FUNCTION_BLOCK "LIOLink_RF200"   // FB5200, SCL
TITLE = LIOLink_RFID / IO_LINK_RFID_1500
{ S7_Optimized_Access := 'FALSE' }
AUTHOR : SIOS
FAMILY : LIOLink
VERSION : 3.0
// IO-Link Device FB for SIMATIC RF200 to use with S7-300/400 controllers! / IO-Link Geraete FB fuer SIMATIC RFID zur Nutzung mit S7-1500!
   VAR_INPUT
      execute : Bool;   // Request to execute function / Auftrag starten (mit steigender Flanke)
      logicalAddr : DInt;   // Logical address of IO-Link master module (sub module for ET 200eco PN) / Logische EA-Adresse des IO-Link Master Moduls
      cap : Int := 227;   // Client Access Point; 0xB400 for ET 200eco PN, CM 8x IO-Link, else 0xE003 (227) / Client Access Point (CAP), Siemens IO-Link Master immer 227 dezimal
      readWrite : Bool;   // FALSE: read, TRUE: write / Lese-/Schreibzugriff: 0=Lesen, 1=Schreiben
      port : Int;   // Port of the IO-Link Master for the Device / Port des Geraetes am IO-Link Mastermodul
      directParameterPage : Bool;   // Read access on parameter page 0 / Lesen Parameter Page 0
      vendorName : Bool;   // Read vendor name / Lesen Herstellername
      vendorText : Bool;   // Read vendor text / Lesen Herstellertext
      productName : Bool;   // Read product name / Lesen Produktname
      productID : Bool;   // Read product ID / Lesen Produkt ID
      fwRevision : Bool;   // Read firmware revision / Lesen FW-Revision
      appSpecificName : Bool;   // Read/write application specific name / Lesen/Schreiben des spezifischen Applikationsnamen
      errorCount : Bool;   // Read number of errors / Lesen des Fehlerzaehlers
      eventHistory : Bool;   // Read event history / Lesen der Ereignishistorie
      readerStatus : Bool;   // Read reader status / Lesen des Reader Status
      tagStatus : Bool;   // Read tag status / Lesen des Variablenstatus
      uidHistory : Bool;   // Read UID history / Lesen des UID Historie
   END_VAR
   VAR_OUTPUT
      done : Bool;   // TRUE: Commanded functionality has been completed successfully / Gueltigkeit 0: Daten ungueltig ; 1: Daten gueltig
      busy : Bool;   // TRUE: FB is not finished and new output values can be expected / 0: Auftrag beendet 1: Auftrag in Bearbeitung
      error : Bool;   // TRUE: An error occurred during the execution of the FB / Fehler = 0: kein Fehler; 1: Funktionsabbruch mit Fehler
      status : Word;   // 16#0000 - 16#7FFF: Status of the FB, 16#8000 - 16#FFFF: Error identification / DP/ PNIO - Fehlerstatus ; ERROR = 1 - Kommunikationsfehler in Detail
      diagDeviceFB : "LIOLink_typeDiagnostics";   // Diagnostics information of LIOLink_Device / IO-Link - Fehlerstatus; ERROR = 1: IO-Link Fehler in Detail
   END_VAR
   VAR_IN_OUT
      data : "LIOLink_RF200_typeAll";   // Data area, device specific (Data Type) / Ablage der Gerätedaten, gerätespezifisch (Datentyp in DB)
   END_VAR
   VAR
      instDevice : "LIOLink_Device";
      statRecordParam : Struct   // Parameters to read/write specific records / Datensatzparameter (geraetespezifisch)
         index : Array[0..28] of Int;   // Index of data set / Datensatzindex
         subindex : Array[0..28] of Int;   // Subindex of data sets / Datensatzsubindex
         length : Array[0..28] of Int;   // Length of data set / Datensatzlänge
      END_STRUCT;
      statRecord : Array[0..231] of Byte;   // Record buffer
      statParameterPage0 AT statRecord : "LIOLink_typeParameterPage0";
      statVendorName AT statRecord : String[12];
      statVendorText AT statRecord : String[12];
      statProductName AT statRecord : String[24];
      statProductID AT statRecord : String[16];
      statFWRevision AT statRecord : String[12];
      statAppSpecName AT statRecord : String[32];
      statErrorCount AT statRecord : Word;
      statEventHistory AT statRecord : "LIOLink_RF200_typeEventHistory";
      statReaderStatus AT statRecord : "LIOLink_RF200_typeReaderStatus";
      statTagStatus AT statRecord : "LIOLink_RF200_typeTagStatus";
      statUIDHistory AT statRecord : "LIOLink_RF200_typeUIDHistory";
      statIndex : Int;   // Requested index
      statSubindex : Int;   // Requested subindex
      statRecordLen : Int;   // Length of record to be written
      statRequest : Int;   // Case of request (data set) / Aktueller Fall (anfgefragter Datensatz)
      statDoneOld : Bool;   // Last cycle's value of instDevice.done
   END_VAR
   VAR_TEMP
      tempIndex : Int;   // Loop index
      tempLen : Int;   // Length
   END_VAR
   VAR CONSTANT
      MODE_READ : Bool := FALSE;   // Mode to read data
      MODE_WRITE : Bool := TRUE;   // Mode to write data
      STATUS_IDLE : Word := 16#7000;   // Status: Idle
   END_VAR
   // statRecordParam.index[0] := 0;
   // statRecordParam.index[1] := 0;
   // statRecordParam.index[2] := 0;
   // statRecordParam.index[3] := 0;
   // statRecordParam.index[4] := 0;
   // statRecordParam.index[5] := 0;
   // statRecordParam.index[6] := 0;
   // statRecordParam.index[7] := 0;
   // statRecordParam.index[8] := 0;
   // statRecordParam.index[9] := 74;
   // statRecordParam.index[10] := 16;
   // statRecordParam.index[11] := 17;
   // statRecordParam.index[12] := 18;
   // statRecordParam.index[13] := 19;
   // statRecordParam.index[14] := 20;
   // statRecordParam.index[15] := 21;
   // statRecordParam.index[16] := 22;
   // statRecordParam.index[17] := 23;
   // statRecordParam.index[18] := 24;
   // statRecordParam.index[19] := 32;
   // statRecordParam.index[20] := 0;
   // statRecordParam.index[21] := 0;
   // statRecordParam.index[22] := 91;
   // statRecordParam.index[23] := 90;
   // statRecordParam.index[24] := 92;
   // statRecordParam.index[25] := 0;
   // statRecordParam.index[26] := 0;
   // statRecordParam.index[27] := 0;
   // statRecordParam.index[28] := 0;
   // statRecordParam.length[0] := 0;
   // statRecordParam.length[1] := 16;
   // statRecordParam.length[2] := 0;
   // statRecordParam.length[3] := 0;
   // statRecordParam.length[4] := 0;
   // statRecordParam.length[5] := 0;
   // statRecordParam.length[6] := 0;
   // statRecordParam.length[7] := 0;
   // statRecordParam.length[8] := 0;
   // statRecordParam.length[9] := 20;
   // statRecordParam.length[10] := 12;
   // statRecordParam.length[11] := 12;
   // statRecordParam.length[12] := 24;
   // statRecordParam.length[13] := 16;
   // statRecordParam.length[14] := 0;
   // statRecordParam.length[15] := 0;
   // statRecordParam.length[16] := 0;
   // statRecordParam.length[17] := 12;
   // statRecordParam.length[18] := 32;
   // statRecordParam.length[19] := 2;
   // statRecordParam.length[20] := 0;
   // statRecordParam.length[21] := 0;
   // statRecordParam.length[22] := 15;
   // statRecordParam.length[23] := 18;
   // statRecordParam.length[24] := 40;
   // statRecordParam.length[25] := 0;
   // statRecordParam.length[26] := 0;
   // statRecordParam.length[27] := 0;
   // statRecordParam.length[28] := 0;
BEGIN
   REGION BLOCK INFO HEADER
     //===============================================================================
     // Siemens / (c)Copyright 2020
     //-------------------------------------------------------------------------------
     // Title:            LIOLink_RF200
     // Function:         Capsule block to communicate with SIMATIC RF200 Readers
     // Library:          LIOLink
     // Author:           Siemens Industry Online Support
     // Tested with:      CPU 317-2 PN/DP FW 3.2
     // Engineering:      TIA Portal V16
     // Restrictions:     --
     // Requirements:     --
     //-------------------------------------------------------------------------------
     // Change log table:
     // Version  | Date       | Expert in charge       | Changes applied
     //----------|------------|------------------------|------------------------------
     // 01.00.00 | 11.04.2014 | Online Support         | First release
     // 02.00.00 | 30.03.2015 | Online Support         | Upgrade to TIA Portal V13 SP1, use function IO_LINK_DEVICE, only one function for S7-1200 and 1500
     // 02.01.00 | 23.10.2015 | Online Support         | Update to IO_LINK_DEVICE Version 3.1
     // 03.00.00 | 22.09.2020 | Online Support         | Upgraded FB "LIOLink_Device" to V4.0.0
     //===============================================================================
   END_REGION

   REGION INIT
     IF (#execute = TRUE AND #instDevice.status = #STATUS_IDLE) THEN
       // Request selector
       IF #directParameterPage THEN
         #statRequest := 1;
       ELSIF #eventHistory THEN
         #statRequest := 9;
       ELSIF #vendorName THEN
         #statRequest := 10;
       ELSIF #vendorText THEN
         #statRequest := 11;
       ELSIF #productName THEN
         #statRequest := 12;
       ELSIF #productID THEN
         #statRequest := 13;
       ELSIF #fwRevision THEN
         #statRequest := 17;
       ELSIF #appSpecificName THEN
         #statRequest := 18;
       ELSIF #errorCount THEN
         #statRequest := 19;
       ELSIF #tagStatus THEN
         #statRequest := 22;
       ELSIF #readerStatus THEN
         #statRequest := 23;
       ELSIF #uidHistory THEN
         #statRequest := 24;
       ELSE
         #statRequest := 0;
       END_IF;

       // Set request specific parameters
       #statIndex := #statRecordParam.index[#statRequest];
       #statSubindex := #statRecordParam.subindex[#statRequest];
       #statRecordLen := #statRecordParam.length[#statRequest];

       IF #readWrite = #MODE_WRITE THEN
         REGION write
           CASE #statRequest OF
             18:
               #statAppSpecName := #data.appSpecificName; // copy text into writing data
               #tempLen := LEN(#statAppSpecName); // determine length of text

               // Shift chars in array to remove String header
               FOR #tempIndex := 0 TO #tempLen - 1 DO
                 #statRecord[#tempIndex] := #statRecord[#tempIndex + 2]; // move [2] to [0], [3] to [1] ... until end of String
               END_FOR;

               // Fill remaining characters with null
               FOR #tempIndex := #tempLen TO #statRecordLen - 1 DO
                 #statRecord[#tempIndex] := CHAR_TO_BYTE('$00');
               END_FOR;
             ELSE // all other data sets are read only  
               ;
           END_CASE;
         END_REGION

       END_IF;
     END_IF;
   END_REGION

   REGION CALL
     #instDevice(execute     := #execute,
                 logicalAddr := #logicalAddr,
                 cap         := #cap,
                 readWrite   := #readWrite,
                 "port"      := #port,
                 index       := #statIndex,
                 subindex    := #statSubindex,
                 writeLen    := #statRecordLen,
                 timeout     := T#20s,
                 record      := #statRecord);
   END_REGION

   REGION READ
     // Copy data if available and valid
     IF #instDevice.done = TRUE AND #statDoneOld = FALSE AND #readWrite = #MODE_READ THEN
       IF (#statRequest >= 10 AND #statRequest <= 18) THEN // Only applies for STRING parameters (case 10..18)
         // add two to data set length for STRING parameters (max./current length)
         FOR #tempIndex := (#statRecordLen + 1) TO 2 BY -1 DO
           #statRecord[#tempIndex] := #statRecord[#tempIndex - 2];
         END_FOR; // Shift chars in array to make space for max/current length of STRING

         #statRecord[0] := INT_TO_BYTE(#statRecordLen); // manipulate array values for STRING 
         #statRecord[1] := INT_TO_BYTE(#statRecordLen);
       END_IF; // Shift all strings and add string header 

       CASE #statRequest OF
         1:
           #data.directParameterPage := #statParameterPage0;
         9:
           #data.eventHistory := #statEventHistory;
         10:
           #data.vendorName := #statVendorName;
         11:
           #data.vendorText := #statVendorText;
         12:
           #data.productName := #statProductName;
         13:
           #data.productID := #statProductID;
         17:
           #data.fwRevision := #statFWRevision;
         18:
           #data.appSpecificName := #statAppSpecName;
         19:
           #data.errorCount := #statErrorCount;
         22:
           #data.tagStatus := #statTagStatus;
         23:
           #data.readerStatus := #statReaderStatus;
         24:
           #data.uidHistory := #statUIDHistory;
         ELSE // Other data sets are not defined
           ;
       END_CASE;
     END_IF;

     #statDoneOld := #instDevice.done;
   END_REGION

   REGION OUTPUTS
     #done := #instDevice.done;
     #busy := #instDevice.busy;
     #error := #instDevice.error;
     #status := #instDevice.status;
     #diagDeviceFB := #instDevice.diagnostics;
   END_REGION
END_FUNCTION_BLOCK

// folder: Device-specific blocks/SIRIUS

FUNCTION_BLOCK "LIOLink_3RA"   // FB5100, SCL
TITLE = LIOLink_3RA / IO_LINK_3RAxy
{ S7_Optimized_Access := 'FALSE' }
AUTHOR : SIOS
FAMILY : LIOLink
VERSION : 3.0
// IO-Link Device FB for SIRIUS 3RAxy to use with S7-300/400 controllers! / IO-Link Geraete FB fuer SIRIUS 3RAxy zur Nutzung mit S7-1500!
   VAR_INPUT
      execute : Bool;   // Request to execute function / Auftrag starten (mit steigender Flanke)
      logicalAddr : DInt;   // Logical address of IO-Link master module (sub module for ET 200eco PN) / Logische EA-Adresse des IO-Link Master Moduls
      cap : Int := 227;   // Client Access Point; 0xB400 for ET 200eco PN, CM 8x IO-Link, else 0xE003 (227) / Client Access Point (CAP), Siemens IO-Link Master immer 227 dezimal
      readWrite : Bool;   // FALSE: read, TRUE: write / Lese-/Schreibzugriff: 0=Lesen, 1=Schreiben
      port : Int;   // Port of the IO-Link Master for the Device / Port des Geraetes am IO-Link Mastermodul
      parameterPage0 : Bool;   // Read access on parameter page 0 / Lesen Parameter Page 0
      parameterPage1 : Bool;   // Read/Write access on parameter page 1 / Lesen-/Schreiben Parameter Page 1
      vendorName : Bool;   // Read Vendor Name / Lesen Herstellername
      vendorText : Bool;   // Read Vendor Text / Lesen Herstellertext
      productName : Bool;   // Read Product Name / Lesen Produktname
      productID : Bool;   // Read Product ID / Lesen Produkt ID
      productText : Bool;   // Read Product Text / Lesen Produkttext
      serialNumber : Bool;   // Read Serial Number / Lesen Seriennummer
      hwRevision : Bool;   // Read HW-Revision / Lesen HW-Revision
      fwRevision : Bool;   // Read FW-Revision / Lesen FW-Revision
      appSpecificName : Bool;   // Read/Write Application Specific Name / Lesen/Schreiben des spezifischen Applikationsnamen
      diagnostics : Bool;   // Read diagnostics / Lesen der Gruppendiagnose
      actualConfig : Bool;   // Read actual configuration / Lesen der Istkonfiguration
      targetConfig : Bool;   // Read/Write target configuration / Lesen/Schreiben der Sollkonfiguration
   END_VAR
   VAR_OUTPUT
      done : Bool;   // TRUE: Commanded functionality has been completed successfully / Gueltigkeit 0: Daten ungueltig ; 1: Daten gueltig
      busy : Bool;   // TRUE: FB is not finished and new output values can be expected / 0: Auftrag beendet 1: Auftrag in Bearbeitung
      error : Bool;   // TRUE: An error occurred during the execution of the FB / Fehler = 0: kein Fehler; 1: Funktionsabbruch mit Fehler
      status : Word;   // 16#0000 - 16#7FFF: Status of the FB, 16#8000 - 16#FFFF: Error identification / DP/ PNIO - Fehlerstatus ; ERROR = 1 - Kommunikationsfehler in Detail
      diagDeviceFB : "LIOLink_typeDiagnostics";   // Diagnostics information of LIOLink_Device / IO-Link - Fehlerstatus; ERROR = 1: IO-Link Fehler in Detail
   END_VAR
   VAR_IN_OUT
      data : "LIOLink_3RA_typeAll";   // Data area, device specific (Data Type) / Ablage der Gerätedaten, gerätespezifisch (Datentyp in DB)
   END_VAR
   VAR
      instDevice : "LIOLink_Device";
      statRecordParam : Struct   // Parameters to read/write specific records / Datensatzparameter (geraetespezifisch)
         index : Array[0..28] of Int;   // Index of data set / Datensatzindex
         subindex : Array[0..28] of Int;   // Subindex of data sets / Datensatzsubindex
         length : Array[0..28] of Int;   // Length of data set / Datensatzlänge
      END_STRUCT;
      statRecord : Array[0..231] of Byte;   // Record buffer
      statParameterPage0 AT statRecord : "LIOLink_typeParameterPage0";
      statVendorName AT statRecord : String[10];
      statVendorText AT statRecord : String[58];
      statProductName AT statRecord : String[30];
      statProductID AT statRecord : String[8];
      statProductText AT statRecord : String[2];
      statSerialNumber AT statRecord : String[8];
      statHWRevision AT statRecord : String[4];
      statFWRevision AT statRecord : String[4];
      statAppSpecName AT statRecord : String[32];
      statDiagnostics AT statRecord : "DIAG_3RAxy";
      statActualConfig AT statRecord : "PARA_3RAxy";
      statTargetConfig AT statRecord : "PARA_3RAxy";
      statParameterPage1 AT statRecord : "ParameterPage1_3RAxy";
      statIndex : Int;   // Requested index
      statSubindex : Int;   // Requested subindex
      statRecordLen : Int;   // Length of record to be written
      statRequest : Int;   // Case of request (data set) / Aktueller Fall (anfgefragter Datensatz)
      statDoneOld : Bool;   // Last cycle's value of instDevice.done
   END_VAR
   VAR_TEMP
      tempIndex : Int;   // Loop index
      tempLen : Int;   // Length
   END_VAR
   VAR CONSTANT
      MODE_READ : Bool := FALSE;   // Mode to read data
      MODE_WRITE : Bool := TRUE;   // Mode to write data
      STATUS_IDLE : Word := 16#7000;   // Status: Idle
   END_VAR
   // statRecordParam.index[4] := 0;
   // statRecordParam.index[3] := 0;
   // statRecordParam.index[2] := 1;
   // statRecordParam.index[1] := 0;
   // statRecordParam.index[25] := 0;
   // statRecordParam.index[24] := 0;
   // statRecordParam.index[23] := 90;
   // statRecordParam.index[21] := 0;
   // statRecordParam.index[20] := 0;
   // statRecordParam.index[18] := 24;
   // statRecordParam.index[17] := 23;
   // statRecordParam.index[16] := 22;
   // statRecordParam.index[15] := 21;
   // statRecordParam.index[14] := 20;
   // statRecordParam.index[13] := 19;
   // statRecordParam.index[12] := 18;
   // statRecordParam.index[11] := 17;
   // statRecordParam.index[10] := 16;
   // statRecordParam.index[8] := 0;
   // statRecordParam.index[7] := 0;
   // statRecordParam.index[6] := 0;
   // statRecordParam.index[5] := 0;
   // statRecordParam.length[28] := 0;
   // statRecordParam.length[27] := 43;
   // statRecordParam.length[26] := 43;
   // statRecordParam.length[25] := 0;
   // statRecordParam.length[24] := 0;
   // statRecordParam.length[23] := 53;
   // statRecordParam.length[22] := 0;
   // statRecordParam.length[21] := 0;
   // statRecordParam.length[20] := 0;
   // statRecordParam.length[19] := 0;
   // statRecordParam.length[18] := 32;
   // statRecordParam.length[17] := 4;
   // statRecordParam.length[16] := 4;
   // statRecordParam.length[15] := 8;
   // statRecordParam.length[14] := 2;
   // statRecordParam.length[13] := 8;
   // statRecordParam.length[12] := 30;
   // statRecordParam.length[11] := 58;
   // statRecordParam.length[10] := 10;
   // statRecordParam.length[9] := 0;
   // statRecordParam.length[8] := 0;
   // statRecordParam.length[7] := 0;
   // statRecordParam.length[6] := 0;
   // statRecordParam.length[5] := 0;
   // statRecordParam.length[4] := 0;
   // statRecordParam.length[3] := 0;
   // statRecordParam.length[2] := 16;
   // statRecordParam.length[1] := 16;
   // statRecordParam.length[0] := 0;
   // statRecordParam.index[28] := 0;
   // statRecordParam.index[27] := 130;
   // statRecordParam.index[26] := 105;
BEGIN
   REGION BLOCK INFO HEADER
     //===============================================================================
     // Siemens / (c)Copyright 2020
     //-------------------------------------------------------------------------------
     // Title:            LIOLink_3RA
     // Function:         Capsule block to communicate with 3RA devices
     // Library:          LIOLink
     // Author:           Siemens Industry Online Support
     // Tested with:      CPU 317-2 PN/DP FW 3.2
     // Engineering:      TIA Portal V16
     // Restrictions:     --
     // Requirements:     --
     //-------------------------------------------------------------------------------
     // Change log table:
     // Version  | Date       | Expert in charge       | Changes applied
     //----------|------------|------------------------|------------------------------
     // 01.00.00 | 11.04.2014 | Online Support         | First release
     // 02.00.00 | 30.03.2015 | Online Support         | Upgrade to TIA Portal V13 SP1, use function IO_LINK_DEVICE, only one function for S7-1200 and 1500
     // 02.01.00 | 23.10.2015 | Online Support         | Update to IO_LINK_DEVICE V3.1.0
     // 03.00.00 | 22.09.2020 | Online Support         | Rewrote block for FB "LIOLink_Device" V4.0.0
     //===============================================================================
   END_REGION

   REGION INIT
     IF (#execute = TRUE AND #instDevice.status = #STATUS_IDLE) THEN
       // Request selector
       IF #parameterPage0 THEN
         #statRequest := 1;
       ELSIF #parameterPage1 THEN
         #statRequest := 2;
       ELSIF #vendorName THEN
         #statRequest := 10;
       ELSIF #vendorText THEN
         #statRequest := 11;
       ELSIF #productName THEN
         #statRequest := 12;
       ELSIF #productID THEN
         #statRequest := 13;
       ELSIF #productText THEN
         #statRequest := 14;
       ELSIF #serialNumber THEN
         #statRequest := 15;
       ELSIF #hwRevision THEN
         #statRequest := 16;
       ELSIF #fwRevision THEN
         #statRequest := 17;
       ELSIF #appSpecificName THEN
         #statRequest := 18;
       ELSIF #diagnostics THEN
         #statRequest := 23;
       ELSIF #actualConfig THEN
         #statRequest := 26;
       ELSIF #targetConfig THEN
         #statRequest := 27;
       ELSE
         #statRequest := 0;
       END_IF;

       #statIndex := #statRecordParam.index[#statRequest];
       #statSubindex := #statRecordParam.subindex[#statRequest];
       #statRecordLen := #statRecordParam.length[#statRequest];

       IF #readWrite = #MODE_WRITE THEN
         REGION write
           CASE #statRequest OF
             2:
               #statParameterPage1 := #data.parameterPage1;
             18:
               #statAppSpecName := #data.appSpecificName; // copy text into writing data
               #tempLen := LEN(#statAppSpecName); // determine length of text

               // Shift chars in array to remove String header
               FOR #tempIndex := 0 TO #tempLen - 1 DO
                 #statRecord[#tempIndex] := #statRecord[#tempIndex + 2]; // move [2] to [0], [3] to [1] ... until end of String
               END_FOR;

               // Fill remaining characters with null
               FOR #tempIndex := #tempLen TO #statRecordLen - 1 DO
                 #statRecord[#tempIndex] := CHAR_TO_BYTE('$00');
               END_FOR;
             27:
               #statTargetConfig := #data.targetConfig;
             ELSE // all other data sets are read only  
               ;
           END_CASE;
         END_REGION

       END_IF;
     END_IF;
   END_REGION

   REGION CALL
     #instDevice(execute     := #execute,
                 logicalAddr := #logicalAddr,
                 cap         := #cap,
                 readWrite   := #readWrite,
                 "port"      := #port,
                 index       := #statIndex,
                 subindex    := #statSubindex,
                 writeLen    := #statRecordLen,
                 timeout     := T#20s,
                 record      := #statRecord);
   END_REGION

   REGION READ
     // Copy data if available and valid
     IF #instDevice.done = TRUE AND #statDoneOld = FALSE AND #readWrite = #MODE_READ THEN
       IF (#statRequest >= 10 AND #statRequest <= 18) THEN // Only applies for STRING parameters (case 10..18)
         // add two to data set length for STRING parameters (max./current length)
         FOR #tempIndex := (#statRecordLen + 1) TO 2 BY -1 DO
           #statRecord[#tempIndex] := #statRecord[#tempIndex - 2];
         END_FOR; // Shift chars in array to make space for max/current length of STRING

         #statRecord[0] := INT_TO_BYTE(#statRecordLen); // manipulate array values for STRING 
         #statRecord[1] := INT_TO_BYTE(#statRecordLen);
       END_IF; // Shift all strings and add string header 

       CASE #statRequest OF
         1:
           #data.parameterPage0 := #statParameterPage0;
         2:
           #data.parameterPage1 := #statParameterPage1;
         10:
           #data.vendorName := #statVendorName;
         11:
           #data.vendorText := #statVendorText;
         12:
           #data.productName := #statProductName;
         13:
           #data.productID := #statProductID;
         14:
           #data.productText := #statProductText;
         15:
           #data.serialNumber := #statSerialNumber;
         16:
           #data.hwRevision := #statHWRevision;
         17:
           #data.fwRevision := #statFWRevision;
         18:
           #data.appSpecificName := #statAppSpecName;
         23:
           #data.diagnostics := #statDiagnostics;
         26:
           #data.actualConfig := #statActualConfig;
         27:
           #data.targetConfig := #statTargetConfig;
         ELSE  // all other data set are not defined
           ;
       END_CASE;
     END_IF;

     #statDoneOld := #instDevice.done;
   END_REGION

   REGION OUTPUTS
     #done := #instDevice.done;
     #busy := #instDevice.busy;
     #error := #instDevice.error;
     #status := #instDevice.status;
     #diagDeviceFB := #instDevice.diagnostics;
   END_REGION
END_FUNCTION_BLOCK

FUNCTION_BLOCK "LIOLink_3RB24"   // FB5110, SCL
TITLE = LIOLink_3RB24 / IO_LINK_3RB24_1500
{ S7_Optimized_Access := 'FALSE' }
AUTHOR : SIOS
FAMILY : LIOLink
VERSION : 3.0
// IO-Link Device FB for SIRIUS 3RB24  to use with S7-300/400 controllers! / IO-Link Geraete FB fuer SIRIUS 3RB24 zur Nutzung mit S7-1500!
   VAR_INPUT
      execute : Bool;   // Request to execute function / Auftrag starten (mit steigender Flanke)
      logicalAddr : DInt;   // Logical address of IO-Link master module (sub module for ET 200eco PN) / Logische EA-Adresse des IO-Link Master Moduls
      cap : Int := 227;   // Client Access Point; 0xB400 for ET 200eco PN, CM 8x IO-Link, else 0xE003 (227) / Client Access Point (CAP), Siemens IO-Link Master immer 227 dezimal
      readWrite : Bool;   // FALSE: read, TRUE: write / Lese-/Schreibzugriff: 0=Lesen, 1=Schreiben
      port : Int;   // Port of the IO-Link Master for the Device / Port des Geraetes am IO-Link Mastermodul
      parameterPage0 : Bool;   // Read access on parameter page 0 / Lesen Parameter Page 0
      vendorName : Bool;   // Read Vendor Name / Lesen Herstellername
      vendorText : Bool;   // Read Vendor Text / Lesen Herstellertext
      productName : Bool;   // Read product name / Lesen Produktname
      productID : Bool;   // Read product ID / Lesen Produkt ID
      productText : Bool;   // Read product text / Lesen Produkttext
      serialNumber : Bool;   // Read serial number / Lesen Seriennummer
      hwRevision : Bool;   // Read hardware revision / Lesen HW-Revision
      fwRevision : Bool;   // Read firmware revision / Lesen FW-Revision
      appSpecificName : Bool;   // Read/Write application specific name / Lesen/Schreiben des spezifischen Applikationsnamen
      processInput : Bool;   // Read process input / Lesen der Prozesseingangsdaten
      processOutput : Bool;   // Read process output / Lesen der Prozesseausgangsdaten
      diagnostics : Bool;   // Read diagnostics / Lesen der Diagnose
      measurements : Bool;   // Read measurements / Lesen der Messwerte
      presetConfigOP : Bool;   // Read/Write preset configuration operator panel / Lesen/Schreiben der Sollkonfiguration Bediengerät
      techFunctions : Bool;   // Read technology functions / Lesen der Technologiefunktionen
   END_VAR
   VAR_OUTPUT
      done : Bool;   // TRUE: Commanded functionality has been completed successfully / Gueltigkeit 0: Daten ungueltig ; 1: Daten gueltig
      busy : Bool;   // TRUE: FB is not finished and new output values can be expected / 0: Auftrag beendet 1: Auftrag in Bearbeitung
      error : Bool;   // TRUE: An error occurred during the execution of the FB / Fehler = 0: kein Fehler; 1: Funktionsabbruch mit Fehler
      status : Word;   // 16#0000 - 16#7FFF: Status of the FB, 16#8000 - 16#FFFF: Error identification / DP/ PNIO - Fehlerstatus ; ERROR = 1 - Kommunikationsfehler in Detail
      diagDeviceFB : "LIOLink_typeDiagnostics";   // Diagnostics information of LIOLink_Device / IO-Link - Fehlerstatus; ERROR = 1: IO-Link Fehler in Detail
   END_VAR
   VAR_IN_OUT
      data : "LIOLink_3RB24_typeAll";   // Data area, device specific (Data Type) / Ablage der Gerätedaten, gerätespezifisch (Datentyp in DB)
   END_VAR
   VAR
      instDevice : "LIOLink_Device";
      statRecordParam : Struct   // Parameters to read/write specific records / Datensatzparameter (geraetespezifisch)
         index : Array[0..28] of Int;   // Index of data set / Datensatzindex
         subindex : Array[0..28] of Int;   // Subindex of data sets / Datensatzsubindex
         length : Array[0..28] of Int;   // Length of data set / Datensatzlänge
      END_STRUCT;
      statRecord : Array[0..231] of Byte;   // Record buffer
      statParameterPage0 AT statRecord : "LIOLink_typeParameterPage0";
      statVendorName AT statRecord : String[10];
      statVendorText AT statRecord : String[64];
      statProductName AT statRecord : String[30];
      statProductID AT statRecord : String[12];
      statProductText AT statRecord : String[2];
      statSerialNumber AT statRecord : String[8];
      statHWRevision AT statRecord : String[4];
      statFWRevision AT statRecord : String[4];
      statAppSpecName AT statRecord : String[32];
      statDiagnostics AT statRecord : "DIAG_3RB24";
      statMeasurements AT statRecord : "MEAS_3RB24";
      statPresetConfigOP AT statRecord : "PresetConfigOP_3RB24";
      statTechFunctions AT statRecord : "TechnoFunctions_3RB24";   // Product family SIRIUS (0x60)
      statProcessInput AT statRecord : Word;
      statProcessOutput AT statRecord : Byte;
      statIndex : Int;   // Requested index
      statSubindex : Int;   // Requested subindex
      statRecordLen : Int;   // Length of record to be written
      statRequest : Int;   // Case of request (data set) / Aktueller Fall (anfgefragter Datensatz)
      statDoneOld : Bool;   // Last cycle's value of instDevice.done
   END_VAR
   VAR_TEMP
      tempIndex : Int;   // Loop index
      tempLen : Int;   // Length
   END_VAR
   VAR CONSTANT
      MODE_READ : Bool := FALSE;   // Mode to read data
      MODE_WRITE : Bool := TRUE;   // Mode to write data
      STATUS_IDLE : Word := 16#7000;   // Status: Idle
   END_VAR
   // statRecordParam.index[4] := 0;
   // statRecordParam.index[3] := 0;
   // statRecordParam.index[2] := 0;
   // statRecordParam.index[1] := 0;
   // statRecordParam.index[25] := 94;
   // statRecordParam.index[24] := 92;
   // statRecordParam.index[23] := 0;
   // statRecordParam.index[21] := 41;
   // statRecordParam.index[20] := 40;
   // statRecordParam.index[18] := 24;
   // statRecordParam.index[17] := 23;
   // statRecordParam.index[16] := 22;
   // statRecordParam.index[15] := 21;
   // statRecordParam.index[14] := 20;
   // statRecordParam.index[13] := 19;
   // statRecordParam.index[12] := 18;
   // statRecordParam.index[11] := 17;
   // statRecordParam.index[6] := 0;
   // statRecordParam.index[5] := 0;
   // statRecordParam.index[10] := 16;
   // statRecordParam.index[8] := 0;
   // statRecordParam.index[7] := 0;
   // statRecordParam.length[28] := 26;
   // statRecordParam.length[27] := 22;
   // statRecordParam.length[26] := 0;
   // statRecordParam.length[25] := 40;
   // statRecordParam.length[24] := 25;
   // statRecordParam.length[23] := 0;
   // statRecordParam.length[22] := 0;
   // statRecordParam.length[21] := 1;
   // statRecordParam.length[20] := 2;
   // statRecordParam.length[19] := 0;
   // statRecordParam.length[18] := 32;
   // statRecordParam.length[17] := 4;
   // statRecordParam.length[16] := 4;
   // statRecordParam.length[15] := 8;
   // statRecordParam.length[14] := 2;
   // statRecordParam.length[13] := 12;
   // statRecordParam.length[12] := 30;
   // statRecordParam.length[11] := 64;
   // statRecordParam.length[10] := 10;
   // statRecordParam.length[9] := 0;
   // statRecordParam.length[8] := 0;
   // statRecordParam.length[7] := 0;
   // statRecordParam.length[6] := 0;
   // statRecordParam.length[5] := 0;
   // statRecordParam.length[4] := 0;
   // statRecordParam.length[3] := 0;
   // statRecordParam.length[2] := 0;
   // statRecordParam.length[1] := 16;
   // statRecordParam.length[0] := 0;
   // statRecordParam.index[28] := 131;
   // statRecordParam.index[27] := 130;
   // statRecordParam.index[26] := 0;
BEGIN
   REGION BLOCK INFO HEADER
     //===============================================================================
     // Siemens / (c)Copyright 2020
     //-------------------------------------------------------------------------------
     // Title:            LIOLink_3RB24
     // Function:         Capsule block to communicate with 3RB24 devices
     // Library:          LIOLink
     // Author:           Siemens Industry Online Support
     // Tested with:      CPU 317-2 PN/DP FW 3.2
     // Engineering:      TIA Portal V16
     // Restrictions:     --
     // Requirements:     --
     //-------------------------------------------------------------------------------
     // Change log table:
     // Version  | Date       | Expert in charge       | Changes applied
     //----------|------------|------------------------|------------------------------
     // 01.00.00 | 11.04.2014 | Online Support         | First release
     // 02.00.00 | 30.03.2015 | Online Support         | Upgrade to TIA Portal V13 SP1, use function IO_LINK_DEVICE, only one function for S7-1200 and 1500
     // 02.01.00 | 23.10.2015 | Online Support         | Update to IO_LINK_DEVICE Version 3.1
     // 03.00.00 | 22.09.2020 | Online Support         | Rewrote block for FB "LIOLink_Device" V4.0.0
     //===============================================================================
   END_REGION

   REGION INIT
     IF (#execute = TRUE AND #instDevice.status = #STATUS_IDLE) THEN
       // Request selector
       IF #parameterPage0 THEN
         #statRequest := 1;
       ELSIF #vendorName THEN
         #statRequest := 10;
       ELSIF #vendorText THEN
         #statRequest := 11;
       ELSIF #productName THEN
         #statRequest := 12;
       ELSIF #productID THEN
         #statRequest := 13;
       ELSIF #productText THEN
         #statRequest := 14;
       ELSIF #serialNumber THEN
         #statRequest := 15;
       ELSIF #hwRevision THEN
         #statRequest := 16;
       ELSIF #fwRevision THEN
         #statRequest := 17;
       ELSIF #appSpecificName THEN
         #statRequest := 18;
       ELSIF #processInput THEN
         #statRequest := 20;
       ELSIF #processOutput THEN
         #statRequest := 21;
       ELSIF #diagnostics THEN
         #statRequest := 24;
       ELSIF #measurements THEN
         #statRequest := 25;
       ELSIF #presetConfigOP THEN
         #statRequest := 27;
       ELSIF #techFunctions THEN
         #statRequest := 28;
       ELSE
         #statRequest := 0;
       END_IF;

       // Set request specific parameters
       #statIndex := #statRecordParam.index[#statRequest];
       #statSubindex := #statRecordParam.subindex[#statRequest];
       #statRecordLen := #statRecordParam.length[#statRequest];

       IF #readWrite = #MODE_WRITE THEN
         REGION write
           CASE #statRequest OF
             18:
               #statAppSpecName := #data.appSpecificName; // copy text into writing data
               #tempLen := LEN(#statAppSpecName); // determine length of text

               // Shift chars in array to remove String header
               FOR #tempIndex := 0 TO #tempLen - 1 DO
                 #statRecord[#tempIndex] := #statRecord[#tempIndex + 2]; // move [2] to [0], [3] to [1] ... until end of String
               END_FOR;

               // Fill remaining characters with null
               FOR #tempIndex := #tempLen TO #statRecordLen - 1 DO
                 #statRecord[#tempIndex] := CHAR_TO_BYTE('$00');
               END_FOR;
             27:
               #statPresetConfigOP := #data.presetConfig;
             ELSE // all other data sets are read only  
               ;
           END_CASE;
         END_REGION

       END_IF;
     END_IF;
   END_REGION

   REGION CALL
     #instDevice(execute     := #execute,
                 logicalAddr := #logicalAddr,
                 cap         := #cap,
                 readWrite   := #readWrite,
                 "port"      := #port,
                 index       := #statIndex,
                 subindex    := #statSubindex,
                 writeLen    := #statRecordLen,
                 timeout     := T#20s,
                 record      := #statRecord);
   END_REGION

   REGION READ
     // Copy data if available and valid
     IF #instDevice.done = TRUE AND #statDoneOld = FALSE AND #readWrite = #MODE_READ THEN
       IF (#statRequest >= 10 AND #statRequest <= 18) THEN // Only applies for STRING parameters (case 10..18)
         // add two to data set length for STRING parameters (max./current length)
         FOR #tempIndex := (#statRecordLen + 1) TO 2 BY -1 DO
           #statRecord[#tempIndex] := #statRecord[#tempIndex - 2];
         END_FOR; // Shift chars in array to make space for max/current length of STRING

         #statRecord[0] := INT_TO_BYTE(#statRecordLen); // manipulate array values for STRING 
         #statRecord[1] := INT_TO_BYTE(#statRecordLen);
       END_IF; // Shift all strings and add string header 

       CASE #statRequest OF
         1:
           #data.parameterPage0 := #statParameterPage0;
         10:
           #data.vendorName := #statVendorName;
         11:
           #data.vendorText := #statVendorText;
         12:
           #data.productName := #statProductName;
         13:
           #data.productID := #statProductID;
         14:
           #data.productText := #statProductText;
         15:
           #data.serialNumber := #statSerialNumber;
         16:
           #data.hwRevision := #statHWRevision;
         17:
           #data.fwRevision := #statFWRevision;
         18:
           #data.appSpecificName := #statAppSpecName;
         20:
           #data.processInput := #statProcessInput;
         21:
           #data.processOutput := #statProcessOutput;
         24:
           #data.diagnostics := #statDiagnostics;
         25:
           #data.measuredValues := #statMeasurements;
         27:
           #data.presetConfig := #statPresetConfigOP;
         28:
           #data.techFunctions := #statTechFunctions;
         ELSE  // Other data sets are not defined
           ;
       END_CASE;
     END_IF;

     #statDoneOld := #instDevice.done;
   END_REGION

   REGION OUTPUTS
     #done := #instDevice.done;
     #busy := #instDevice.busy;
     #error := #instDevice.error;
     #status := #instDevice.status;
     #diagDeviceFB := #instDevice.diagnostics;
   END_REGION
END_FUNCTION_BLOCK

FUNCTION_BLOCK "LIOLink_3RR24"   // FB5120, SCL
TITLE = LIOLink_3RR24 / IO_LINK_3RR24_1500
{ S7_Optimized_Access := 'FALSE' }
AUTHOR : SIOS
FAMILY : LIOLink
VERSION : 3.0
// IO-Link Device FB for SIRIUS 3RR24 to use with S7-300/400 controllers! / IO-Link Geraete FB fuer SIRIUS 3RR24 zur Nutzung mit S7-1500!
   VAR_INPUT
      execute : Bool;   // Request to execute function / Auftrag starten (mit steigender Flanke)
      logicalAddr : DInt;   // Logical address of IO-Link master module (sub module for ET 200eco PN) / Logische EA-Adresse des IO-Link Master Moduls
      cap : Int := 227;   // Client Access Point; 0xB400 for ET 200eco PN, CM 8x IO-Link, else 0xE003 (227) / Client Access Point (CAP), Siemens IO-Link Master immer 227 dezimal
      readWrite : Bool;   // FALSE: read, TRUE: write / Lese-/Schreibzugriff: 0=Lesen, 1=Schreiben
      port : Int;   // Port of the IO-Link Master for the Device / Port des Geraetes am IO-Link Mastermodul
      parameterPage0 : Bool;   // Read access on parameter page 0 / Lesen Parameter Page 0
      systemCommands : Bool;   // Write system commands / Schreiben Systemkommandos
      vendorName : Bool;   // Read vendor name / Lesen Herstellername
      vendorText : Bool;   // Read vendor text / Lesen Herstellertext
      productName : Bool;   // Read product name / Lesen Produktname
      productID : Bool;   // Read product ID / Lesen Produkt ID
      serialNumber : Bool;   // Read serial number / Lesen Seriennummer
      hwRevision : Bool;   // Read hardware revision / Lesen HW-Revision
      fwRevision : Bool;   // Read firmware revision / Lesen FW-Revision
      appSpecificName : Bool;   // Read/Write application specific name / Lesen/Schreiben des spezifischen Applikationsnamen
      diagnostics : Bool;   // Read diagnostics / Lesen der Diagnose
      measurements : Bool;   // Read measurements / Lesen der Messwerte
      parameters : Bool;   // Read/Write parameters / Lesen/Schreiben der Parameter
   END_VAR
   VAR_OUTPUT
      done : Bool;   // TRUE: Commanded functionality has been completed successfully / Gueltigkeit 0: Daten ungueltig ; 1: Daten gueltig
      busy : Bool;   // TRUE: FB is not finished and new output values can be expected / 0: Auftrag beendet 1: Auftrag in Bearbeitung
      error : Bool;   // TRUE: An error occurred during the execution of the FB / Fehler = 0: kein Fehler; 1: Funktionsabbruch mit Fehler
      status : Word;   // 16#0000 - 16#7FFF: Status of the FB, 16#8000 - 16#FFFF: Error identification / DP/ PNIO - Fehlerstatus ; ERROR = 1 - Kommunikationsfehler in Detail
      diagDeviceFB : "LIOLink_typeDiagnostics";   // Diagnostics information of LIOLink_Device / IO-Link - Fehlerstatus; ERROR = 1: IO-Link Fehler in Detail
   END_VAR
   VAR_IN_OUT
      data : "LIOLink_3RR24_typeAll";   // Data area, device specific (Data Type) / Ablage der Gerätedaten, gerätespezifisch (Datentyp in DB)
   END_VAR
   VAR
      instDevice : "LIOLink_Device";
      statRecordParam : Struct   // Parameters to read/write specific records / Datensatzparameter (geraetespezifisch)
         index : Array[0..28] of Int;   // Index of data set / Datensatzindex
         subindex : Array[0..28] of Int;   // Subindex of data sets / Datensatzsubindex
         length : Array[0..28] of Int;   // Length of data set / Datensatzlänge
      END_STRUCT;
      statRecord : Array[0..231] of Byte;   // Record buffer
      statParameterPage0 AT statRecord : "LIOLink_typeParameterPage0";
      statVendorName AT statRecord : String[11];
      statVendorText AT statRecord : String[64];
      statProductName AT statRecord : String[64];
      statProductID AT statRecord : String[14];
      statSerialNumber AT statRecord : String[16];
      statHWRevision AT statRecord : String[7];
      statFWRevision AT statRecord : String[7];
      statAppSpecName AT statRecord : String[32];
      statDiagnostics AT statRecord : "DIAG_3RR24";
      statMeasurements AT statRecord : "MEAS_3RR24";
      statParameters AT statRecord : "PARA_3RR24";   // Product family SIRIUS (0x60)
      statSystemCommands AT statRecord : Byte;
      statIndex : Int;   // Requested index
      statSubindex : Int;   // Requested subindex
      statRecordLen : Int;   // Length of record to be written
      statRequest : Int;   // Case of request (data set) / Aktueller Fall (anfgefragter Datensatz)
      statDoneOld : Bool;   // Last cycle's value of instDevice.done
   END_VAR
   VAR_TEMP
      tempIndex : Int;   // Loop index
      tempLen : Int;   // Length
   END_VAR
   VAR CONSTANT
      MODE_READ : Bool := FALSE;   // Mode to read data
      MODE_WRITE : Bool := TRUE;   // Mode to write data
      STATUS_IDLE : Word := 16#7000;   // Status: Idle
   END_VAR
   // statRecordParam.index[3] := 2;
   // statRecordParam.index[2] := 0;
   // statRecordParam.index[1] := 0;
   // statRecordParam.index[0] := 0;
   // statRecordParam.index[18] := 24;
   // statRecordParam.index[17] := 23;
   // statRecordParam.index[5] := 0;
   // statRecordParam.index[4] := 0;
   // statRecordParam.index[16] := 22;
   // statRecordParam.index[15] := 21;
   // statRecordParam.index[14] := 20;
   // statRecordParam.index[13] := 19;
   // statRecordParam.index[12] := 18;
   // statRecordParam.index[11] := 17;
   // statRecordParam.index[10] := 16;
   // statRecordParam.index[9] := 0;
   // statRecordParam.index[8] := 0;
   // statRecordParam.index[7] := 0;
   // statRecordParam.index[6] := 0;
   // statRecordParam.length[28] := 62;
   // statRecordParam.length[27] := 0;
   // statRecordParam.length[26] := 0;
   // statRecordParam.length[25] := 56;
   // statRecordParam.length[24] := 30;
   // statRecordParam.length[23] := 0;
   // statRecordParam.length[22] := 0;
   // statRecordParam.length[21] := 0;
   // statRecordParam.length[20] := 0;
   // statRecordParam.length[19] := 0;
   // statRecordParam.length[18] := 32;
   // statRecordParam.length[17] := 7;
   // statRecordParam.length[16] := 7;
   // statRecordParam.length[15] := 16;
   // statRecordParam.length[14] := 0;
   // statRecordParam.length[13] := 14;
   // statRecordParam.length[12] := 64;
   // statRecordParam.length[11] := 64;
   // statRecordParam.length[10] := 11;
   // statRecordParam.length[9] := 0;
   // statRecordParam.length[8] := 0;
   // statRecordParam.length[7] := 0;
   // statRecordParam.length[6] := 0;
   // statRecordParam.length[5] := 0;
   // statRecordParam.length[4] := 0;
   // statRecordParam.length[3] := 1;
   // statRecordParam.length[2] := 0;
   // statRecordParam.length[1] := 16;
   // statRecordParam.length[0] := 0;
   // statRecordParam.index[28] := 131;
   // statRecordParam.index[27] := 0;
   // statRecordParam.index[26] := 0;
   // statRecordParam.index[25] := 94;
   // statRecordParam.index[24] := 92;
   // statRecordParam.index[23] := 0;
   // statRecordParam.index[22] := 0;
   // statRecordParam.index[21] := 0;
   // statRecordParam.index[20] := 0;
   // statRecordParam.index[19] := 0;
BEGIN
   REGION BLOCK INFO HEADER
     //===============================================================================
     // Siemens / (c)Copyright 2020
     //-------------------------------------------------------------------------------
     // Title:            LIOLink_3RR24
     // Function:         Capsule block to communicate with 3RR24 devices
     // Library:          LIOLink
     // Author:           Siemens Industry Online Support
     // Tested with:      CPU 317-2 PN/DP FW 3.2
     // Engineering:      TIA Portal V16
     // Restrictions:     --
     // Requirements:     --
     //-------------------------------------------------------------------------------
     // Change log table:
     // Version  | Date       | Expert in charge       | Changes applied
     //----------|------------|------------------------|------------------------------
     // 01.00.00 | 11.04.2014 | Online Support         | First release
     // 01.00.01 | 12.09.2014 | Online Support         | Bugfixing write case 28 (data set 131)
     // 02.00.00 | 30.03.2015 | Online Support         | Upgrade to TIA Portal V13 SP1, use function IO_LINK_DEVICE, only one function for S7-1200 and 1500
     // 02.01.00 | 23.10.2015 | Online Support         | Update to IO_LINK_DEVICE Version 3.1
     // 03.00.00 | 22.09.2020 | Online Support         | Rewrote block for FB "LIOLink_Device" V4.0.0
     //===============================================================================
   END_REGION

   REGION INIT
     IF (#execute = TRUE AND #instDevice.status = #STATUS_IDLE) THEN
       // Request selector
       IF #parameterPage0 THEN
         #statRequest := 1;
       ELSIF #systemCommands THEN
         #statRequest := 3;
       ELSIF #vendorName THEN
         #statRequest := 10;
       ELSIF #vendorText THEN
         #statRequest := 11;
       ELSIF #productName THEN
         #statRequest := 12;
       ELSIF #productID THEN
         #statRequest := 13;
       ELSIF #serialNumber THEN
         #statRequest := 15;
       ELSIF #hwRevision THEN
         #statRequest := 16;
       ELSIF #fwRevision THEN
         #statRequest := 17;
       ELSIF #appSpecificName THEN
         #statRequest := 18;
       ELSIF #diagnostics THEN
         #statRequest := 24;
       ELSIF #measurements THEN
         #statRequest := 25;
       ELSIF #parameters THEN
         #statRequest := 28;
       ELSE
         #statRequest := 0;
       END_IF;

       // Set request specific parameters
       #statIndex := #statRecordParam.index[#statRequest];
       #statSubindex := #statRecordParam.subindex[#statRequest];
       #statRecordLen := #statRecordParam.length[#statRequest];

       IF #readWrite = #MODE_WRITE THEN
         REGION write
           CASE #statRequest OF
             3:
               #statSystemCommands := #data.systemCommands;
             18:
               #statAppSpecName := #data.appSpecificName; // copy text into writing data
               #tempLen := LEN(#statAppSpecName); // determine length of text

               // Shift chars in array to remove String header
               FOR #tempIndex := 0 TO #tempLen - 1 DO
                 #statRecord[#tempIndex] := #statRecord[#tempIndex + 2]; // move [2] to [0], [3] to [1] ... until end of String
               END_FOR;

               // Fill remaining characters with null
               FOR #tempIndex := #tempLen TO #statRecordLen - 1 DO
                 #statRecord[#tempIndex] := CHAR_TO_BYTE('$00');
               END_FOR;
             28:
               #statParameters := #data.parameters;
             ELSE    // all other data set are read only
               ;
           END_CASE;
         END_REGION

       END_IF;
     END_IF;
   END_REGION

   REGION CALL
     #instDevice(execute     := #execute,
                 logicalAddr := #logicalAddr,
                 cap         := #cap,
                 readWrite   := #readWrite,
                 "port"      := #port,
                 index       := #statIndex,
                 subindex    := #statSubindex,
                 writeLen    := #statRecordLen,
                 timeout     := T#20s,
                 record      := #statRecord);
   END_REGION

   REGION READ
     // Copy data if available and valid
     IF #instDevice.done = TRUE AND #statDoneOld = FALSE AND #readWrite = #MODE_READ THEN
       IF (#statRequest >= 10 AND #statRequest <= 18) THEN // Only applies for STRING parameters (case 10..18)
         // add two to data set length for STRING parameters (max./current length)
         FOR #tempIndex := (#statRecordLen + 1) TO 2 BY -1 DO
           #statRecord[#tempIndex] := #statRecord[#tempIndex - 2];
         END_FOR; // Shift chars in array to make space for max/current length of STRING

         #statRecord[0] := INT_TO_BYTE(#statRecordLen); // manipulate array values for STRING 
         #statRecord[1] := INT_TO_BYTE(#statRecordLen);
       END_IF; // Shift all strings and add string header 

       CASE #statRequest OF
         1:
           #data.parameterPage0 := #statParameterPage0;
         10:
           #data.vendorName := #statVendorName;
         11:
           #data.vendorText := #statVendorText;
         12:
           #data.productName := #statProductName;
         13:
           #data.productID := #statProductID;
         15:
           #data.serialNumber := #statSerialNumber;
         16:
           #data.hwRevision := #statHWRevision;
         17:
           #data.fwRevision := #statFWRevision;
         18:
           #data.appSpecificName := #statAppSpecName;
         24:
           #data.diagnostics := #statDiagnostics;
         25:
           #data.measuredValues := #statMeasurements;
         28:
           #data.parameters := #statParameters;
         ELSE  // Other data sets are not defined
           ;
       END_CASE;
     END_IF;

     #statDoneOld := #instDevice.done;
   END_REGION

   REGION OUTPUTS
     #done := #instDevice.done;
     #busy := #instDevice.busy;
     #error := #instDevice.error;
     #status := #instDevice.status;
     #diagDeviceFB := #instDevice.diagnostics;
   END_REGION
END_FUNCTION_BLOCK

FUNCTION_BLOCK "LIOLink_3RS1"   // FB5130, SCL
TITLE = LIOLink_3RS1 / IO_LINK_3RS1x_1500
{ S7_Optimized_Access := 'FALSE' }
AUTHOR : SIOS
FAMILY : LIOLink
VERSION : 3.0
// Capsule block to communicate with SIRIUS 3RS1 devices with S7-300/400 Controllers / IO-Link Geraete FB fuer SIRIUS 3RS1x zur Nutzung mit S7-1500!
   VAR_INPUT
      execute : Bool;   // Request to execute function / Auftrag starten (mit steigender Flanke)
      logicalAddr : DInt;   // Logical address of IO-Link master module (sub module for ET 200eco PN) / Logische EA-Adresse des IO-Link Master Moduls
      cap : Int := 227;   // Client Access Point; 0xB400 for ET 200eco PN, CM 8x IO-Link, else 0xE003 (227) / Client Access Point (CAP), Siemens IO-Link Master immer 227 dezimal
      readWrite : Bool;   // FALSE: read, TRUE: write / Lese-/Schreibzugriff: 0=Lesen, 1=Schreiben
      port : Int;   // Port of the IO-Link Master for the Device / Port des Geraetes am IO-Link Mastermodul
      parameterPage0 : Bool;   // Read access on parameter page 0 / Lesen Parameter Page 0
      vendorName : Bool;   // Read vendor name / Lesen Herstellername
      vendorText : Bool;   // Read vendor text / Lesen Herstellertext
      productName : Bool;   // Read product name / Lesen Produktname
      productID : Bool;   // Read product ID / Lesen Produkt ID
      hwRevision : Bool;   // Read hardware revision / Lesen HW-Revision
      fwRevision : Bool;   // Read firmware revision / Lesen FW-Revision
      appSpecificName : Bool;   // Read/Write application specific name / Lesen/Schreiben des spezifischen Applikationsnamen
      diagnostics : Bool;   // Read diagnostics / Lesen der Diagnose
      measurements : Bool;   // Read measurements / Lesen der Messwerte
      parameters : Bool;   // Read/Write parameters / Lesen/Schreiben der Parameter
   END_VAR
   VAR_OUTPUT
      done : Bool;   // TRUE: Commanded functionality has been completed successfully / Gueltigkeit 0: Daten ungueltig ; 1: Daten gueltig
      busy : Bool;   // TRUE: FB is not finished and new output values can be expected / 0: Auftrag beendet 1: Auftrag in Bearbeitung
      error : Bool;   // TRUE: An error occurred during the execution of the FB / Fehler = 0: kein Fehler; 1: Funktionsabbruch mit Fehler
      status : Word;   // 16#0000 - 16#7FFF: Status of the FB, 16#8000 - 16#FFFF: Error identification / DP/ PNIO - Fehlerstatus ; ERROR = 1 - Kommunikationsfehler in Detail
      diagDeviceFB : "LIOLink_typeDiagnostics";   // Diagnostics information of LIOLink_Device / IO-Link - Fehlerstatus; ERROR = 1: IO-Link Fehler in Detail
   END_VAR
   VAR_IN_OUT
      data : "LIOLink_3RS1_typeAll";   // Data area, device specific (Data Type) / Ablage der Gerätedaten, gerätespezifisch (Datentyp in DB)
   END_VAR
   VAR
      instDevice : "LIOLink_Device";
      statRecordParam : Struct   // Parameters to read/write specific records / Datensatzparameter (geraetespezifisch)
         index : Array[0..28] of Int;   // Index of data set / Datensatzindex
         subindex : Array[0..28] of Int;   // Subindex of data sets / Datensatzsubindex
         length : Array[0..28] of Int;   // Length of data set / Datensatzlänge
      END_STRUCT;
      statRecord : Array[0..231] of Byte;   // Record buffer
      statParameterPage0 AT statRecord : "LIOLink_typeParameterPage0";
      statVendorName AT statRecord : String[11];
      statVendorText AT statRecord : String[64];
      statProductName AT statRecord : String[64];
      statProductID AT statRecord : String[14];
      statHWRevision AT statRecord : String[7];
      statFWRevision AT statRecord : String[7];
      statAppSpecName AT statRecord : String[32];
      statDiagnostics AT statRecord : "DIAG_3RS1x";
      statMeasurements AT statRecord : "MEAS_3RS1x";
      statParameters AT statRecord : "PARA_3RS1x";   // Product family SIRIUS (0x60)
      statIndex : Int;   // Requested index
      statSubindex : Int;   // Requested subindex
      statRecordLen : Int;   // Length of record to be written
      statRequest : Int;   // Case of request (data set) / Aktueller Fall (anfgefragter Datensatz)
      statDoneOld : Bool;   // Last cycle's value of instDevice.done
   END_VAR
   VAR_TEMP
      tempIndex : Int;   // Loop index
      tempLen : Int;   // Length
   END_VAR
   VAR CONSTANT
      MODE_READ : Bool := FALSE;   // Mode to read data
      MODE_WRITE : Bool := TRUE;   // Mode to write data
      STATUS_IDLE : Word := 16#7000;   // Status: Idle
   END_VAR
   // statRecordParam.index[3] := 0;
   // statRecordParam.index[2] := 0;
   // statRecordParam.index[1] := 0;
   // statRecordParam.index[0] := 0;
   // statRecordParam.index[17] := 23;
   // statRecordParam.index[16] := 22;
   // statRecordParam.index[5] := 0;
   // statRecordParam.index[4] := 0;
   // statRecordParam.index[15] := 21;
   // statRecordParam.index[14] := 20;
   // statRecordParam.index[13] := 19;
   // statRecordParam.index[12] := 18;
   // statRecordParam.index[11] := 17;
   // statRecordParam.index[10] := 16;
   // statRecordParam.index[9] := 0;
   // statRecordParam.index[8] := 0;
   // statRecordParam.index[7] := 0;
   // statRecordParam.index[6] := 0;
   // statRecordParam.length[28] := 50;
   // statRecordParam.length[27] := 0;
   // statRecordParam.length[26] := 0;
   // statRecordParam.length[25] := 46;
   // statRecordParam.length[24] := 40;
   // statRecordParam.length[23] := 0;
   // statRecordParam.length[22] := 0;
   // statRecordParam.length[21] := 0;
   // statRecordParam.length[20] := 0;
   // statRecordParam.length[19] := 0;
   // statRecordParam.length[18] := 32;
   // statRecordParam.length[17] := 7;
   // statRecordParam.length[16] := 7;
   // statRecordParam.length[15] := 0;
   // statRecordParam.length[14] := 0;
   // statRecordParam.length[13] := 14;
   // statRecordParam.length[12] := 64;
   // statRecordParam.length[11] := 64;
   // statRecordParam.length[10] := 11;
   // statRecordParam.length[9] := 0;
   // statRecordParam.length[8] := 0;
   // statRecordParam.length[7] := 0;
   // statRecordParam.length[6] := 0;
   // statRecordParam.length[5] := 0;
   // statRecordParam.length[4] := 0;
   // statRecordParam.length[3] := 0;
   // statRecordParam.length[2] := 0;
   // statRecordParam.length[1] := 16;
   // statRecordParam.length[0] := 0;
   // statRecordParam.index[28] := 131;
   // statRecordParam.index[27] := 0;
   // statRecordParam.index[26] := 0;
   // statRecordParam.index[25] := 94;
   // statRecordParam.index[24] := 92;
   // statRecordParam.index[23] := 0;
   // statRecordParam.index[22] := 0;
   // statRecordParam.index[21] := 0;
   // statRecordParam.index[20] := 0;
   // statRecordParam.index[19] := 0;
   // statRecordParam.index[18] := 24;
BEGIN
   REGION BLOCK INFO HEADER
     //===============================================================================
     // Siemens / (c)Copyright 2020
     //-------------------------------------------------------------------------------
     // Title:            LIOLink_3RS1
     // Function:         Capsule block to communicate with SIRIUS 3RS1 devices
     // Library:          LIOLink
     // Author:           Siemens Industry Online Support
     // Tested with:      CPU 317-2 PN/DP FW 3.2
     // Engineering:      TIA Portal V16
     // Restrictions:     --
     // Requirements:     --
     //-------------------------------------------------------------------------------
     // Change log table:
     // Version  | Date       | Expert in charge       | Changes applied
     //----------|------------|------------------------|------------------------------
     // 01.00.00 | 11.04.2014 | Online Support         | First release
     // 02.00.00 | 30.03.2015 | Online Support         | Upgrade to TIA Portal V13 SP1, use function IO_LINK_DEVICE, only one function for S7-1200 and 1500
     // 02.01.00 | 23.10.2015 | Online Support         | Update to IO_LINK_DEVICE Version 3.1
     // 03.00.00 | 22.09.2020 | Online Support         | Rewrote block for FB "LIOLink_Device" V4.0.0
     //===============================================================================
   END_REGION

   REGION INIT
     IF (#execute = TRUE AND #instDevice.status = #STATUS_IDLE) THEN
       // Request selector
       IF #parameterPage0 THEN
         #statRequest := 1;
       ELSIF #vendorName THEN
         #statRequest := 10;
       ELSIF #vendorText THEN
         #statRequest := 11;
       ELSIF #productName THEN
         #statRequest := 12;
       ELSIF #productID THEN
         #statRequest := 13;
       ELSIF #hwRevision THEN
         #statRequest := 16;
       ELSIF #fwRevision THEN
         #statRequest := 17;
       ELSIF #appSpecificName THEN
         #statRequest := 18;
       ELSIF #diagnostics THEN
         #statRequest := 24;
       ELSIF #measurements THEN
         #statRequest := 25;
       ELSIF #parameters THEN
         #statRequest := 28;
       ELSE
         #statRequest := 0;
       END_IF;

       // Set request specific parameters
       #statIndex := #statRecordParam.index[#statRequest];
       #statSubindex := #statRecordParam.subindex[#statRequest];
       #statRecordLen := #statRecordParam.length[#statRequest];

       IF #readWrite = #MODE_WRITE THEN
         REGION write
           CASE #statRequest OF
             18:
               #statAppSpecName := #data.appSpecificName; // copy text into writing data
               #tempLen := LEN(#statAppSpecName); // determine length of text

               // Shift chars in array to remove String header
               FOR #tempIndex := 0 TO #tempLen - 1 DO
                 #statRecord[#tempIndex] := #statRecord[#tempIndex + 2]; // move [2] to [0], [3] to [1] ... until end of String
               END_FOR;

               // Fill remaining characters with null
               FOR #tempIndex := #tempLen TO #statRecordLen - 1 DO
                 #statRecord[#tempIndex] := CHAR_TO_BYTE('$00');
               END_FOR;
             28:
               #statParameters := #data.parameters;
             ELSE // All other data sets are read only
               ;
           END_CASE;
         END_REGION

       END_IF;
     END_IF;
   END_REGION

   REGION CALL
     #instDevice(execute     := #execute,
                 logicalAddr := #logicalAddr,
                 cap         := #cap,
                 readWrite   := #readWrite,
                 "port"      := #port,
                 index       := #statIndex,
                 subindex    := #statSubindex,
                 writeLen    := #statRecordLen,
                 timeout     := T#20s,
                 record      := #statRecord);
   END_REGION

   REGION READ
     // Copy data if available and valid
     IF #instDevice.done = TRUE AND #statDoneOld = FALSE AND #readWrite = #MODE_READ THEN
       IF (#statRequest >= 10 AND #statRequest <= 18) THEN // Only applies for STRING parameters (case 10..18)
         // add two to data set length for STRING parameters (max./current length)
         FOR #tempIndex := (#statRecordLen + 1) TO 2 BY -1 DO
           #statRecord[#tempIndex] := #statRecord[#tempIndex - 2];
         END_FOR; // Shift chars in array to make space for max/current length of STRING

         #statRecord[0] := INT_TO_BYTE(#statRecordLen); // manipulate array values for STRING 
         #statRecord[1] := INT_TO_BYTE(#statRecordLen);
       END_IF; // Shift all strings and add string header 

       CASE #statRequest OF
         1:
           #data.parameterPage0 := #statParameterPage0;
         10:
           #data.vendorName := #statVendorName;
         11:
           #data.vendorText := #statVendorText;
         12:
           #data.productName := #statProductName;
         13:
           #data.productID := #statProductID;
         16:
           #data.hardwareRevision := #statHWRevision;
         17:
           #data.firmwareRevision := #statFWRevision;
         18:
           #data.appSpecificName := #statAppSpecName;
         24:
           #data.diagnostics := #statDiagnostics;
         25:
           #data.measuredValues := #statMeasurements;
         28:
           #data.parameters := #statParameters;
         ELSE  // Other data sets are not defined
           ;
       END_CASE;
     END_IF;

     #statDoneOld := #instDevice.done;
   END_REGION

   REGION OUTPUTS
     #done := #instDevice.done;
     #busy := #instDevice.busy;
     #error := #instDevice.error;
     #status := #instDevice.status;
     #diagDeviceFB := #instDevice.diagnostics;
   END_REGION
END_FUNCTION_BLOCK

FUNCTION_BLOCK "LIOLink_3RS2"   // FB5131, SCL
TITLE = LIOLink_3RS2 / IO_LINK_3RS1x_1500
{ S7_Optimized_Access := 'FALSE' }
AUTHOR : SIOS
FAMILY : LIOLink
VERSION : 1.0
// Capsule block to communicate with SIRIUS 3RS2 devices with S7-300/400 Controllers / IO-Link Geraete FB fuer SIRIUS 3RS1x zur Nutzung mit S7-1500!
   VAR_INPUT
      execute : Bool;   // Request to execute function / Auftrag starten (mit steigender Flanke)
      logicalAddr : DInt;   // Logical address of IO-Link master module (sub module for ET 200eco PN) / Logische EA-Adresse des IO-Link Master Moduls
      cap : Int := 227;   // Client Access Point; 0xB400 for ET 200eco PN, CM 8x IO-Link, else 0xE003 (227) / Client Access Point (CAP), Siemens IO-Link Master immer 227 dezimal
      readWrite : Bool;   // FALSE: read, TRUE: write / Lese-/Schreibzugriff: 0=Lesen, 1=Schreiben
      port : Int;   // Port of the IO-Link Master for the Device / Port des Geraetes am IO-Link Mastermodul
      parameterPage0 : Bool;   // Read parameter page 0 / Lesen Parameter Page 0
      vendorName : Bool;   // Read vendor name / Lesen Herstellername
      vendorText : Bool;   // Read vendor text / Lesen Herstellertext
      productName : Bool;   // Read product name / Lesen Produktname
      productID : Bool;   // Read product ID / Lesen Produkt ID
      fwRevision : Bool;   // Read firmware revision / Lesen FW-Revision
      appSpecificName : Bool;   // Read/write application specific name / Lesen/Schreiben des spezifischen Applikationsnamen
      diagnostics : Bool;   // Read diagnostics / Lesen der Diagnose
      measuredValues : Bool;   // Read measured values / Lesen der Messwerte
      parameters : Bool;   // Read/Write parameters / Lesen/Schreiben der Parameter
   END_VAR
   VAR_OUTPUT
      done : Bool;   // TRUE: Commanded functionality has been completed successfully / Gueltigkeit 0: Daten ungueltig ; 1: Daten gueltig
      busy : Bool;   // TRUE: FB is not finished and new output values can be expected / 0: Auftrag beendet 1: Auftrag in Bearbeitung
      error : Bool;   // TRUE: An error occurred during the execution of the FB / Fehler = 0: kein Fehler; 1: Funktionsabbruch mit Fehler
      status : Word;   // 16#0000 - 16#7FFF: Status of the FB, 16#8000 - 16#FFFF: Error identification / DP/ PNIO - Fehlerstatus ; ERROR = 1 - Kommunikationsfehler in Detail
      diagDeviceFB : "LIOLink_typeDiagnostics";   // Diagnostics information of LIOLink_Device / IO-Link - Fehlerstatus; ERROR = 1: IO-Link Fehler in Detail
   END_VAR
   VAR_IN_OUT
      data : "LIOLink_3RS2_typeAll";   // Data area, device specific (Data Type) / Ablage der Gerätedaten, gerätespezifisch (Datentyp in DB)
   END_VAR
   VAR
      instDevice : "LIOLink_Device";
      statRecord : Array[0..231] of Byte;   // Record buffer
      statParameterPage0 AT statRecord : "LIOLink_typeParameterPage0";
      statVendorName AT statRecord : String[11];
      statVendorText AT statRecord : String[64];
      statProductName AT statRecord : String[64];
      statProductID AT statRecord : String[14];
      statFWRevision AT statRecord : String[7];
      statAppSpecName AT statRecord : String[32];
      statDiagnostics AT statRecord : "LIOLink_3RS2_typeDiag";
      statMeasuredValues AT statRecord : "LIOLink_3RS2_typeMeasure";
      statParameters AT statRecord : "LIOLink_3RS2_typeParam";   // Product family SIRIUS (0x60)
      statIndex : Int;   // Requested index
      statSubindex : Int;   // Requested subindex
      statRecordLen : Int;   // Length of record to be written
      statDoneOld : Bool;   // Last cycle's value of instDevice.done
   END_VAR
   VAR_TEMP
      tempIndex : Int;   // Loop index
      tempLen : Int;   // Length
   END_VAR
   VAR CONSTANT
      MODE_READ : Bool := FALSE;   // Mode to read data
      MODE_WRITE : Bool := TRUE;   // Mode to write data
      STATUS_IDLE : Word := 16#7000;   // Status: Idle
   END_VAR
BEGIN
   REGION BLOCK INFO HEADER
     //===============================================================================
     // Siemens / (c)Copyright 2020
     //-------------------------------------------------------------------------------
     // Title:            LIOLink_3RS2
     // Function:         Capsule block to communicate with SIRIUS 3RS2 devices
     // Library:          LIOLink
     // Author:           Siemens Industry Online Support
     // Tested with:      CPU 317-2 PN/DP FW 3.2
     // Engineering:      TIA Portal V16
     // Restrictions:     --
     // Requirements:     --
     //-------------------------------------------------------------------------------
     // Change log table:
     // Version  | Date       | Expert in charge       | Changes applied
     //----------|------------|------------------------|------------------------------
     // 01.00.00 | 22.09.2020 | Online Support         | First release
     //===============================================================================
   END_REGION

   REGION INIT
     IF (#execute = TRUE AND #instDevice.status = #STATUS_IDLE) THEN
       // Set request-specific parameters
       IF #parameterPage0 THEN
         #statIndex := 0;
         #statRecordLen := 16;
       ELSIF #vendorName THEN
         #statIndex := 16;
         #statRecordLen := 11;
       ELSIF #vendorText THEN
         #statIndex := 17;
         #statRecordLen := 64;
       ELSIF #productName THEN
         #statIndex := 18;
         #statRecordLen := 64;
       ELSIF #productID THEN
         #statIndex := 19;
         #statRecordLen := 14;
       ELSIF #fwRevision THEN
         #statIndex := 23;
         #statRecordLen := 7;
       ELSIF #appSpecificName THEN
         #statIndex := 24;
         #statRecordLen := 32;
       ELSIF #diagnostics THEN
         #statIndex := 92;
         #statRecordLen := 43;
       ELSIF #measuredValues THEN
         #statIndex := 94;
         #statRecordLen := 42;
       ELSIF #parameters THEN
         #statIndex := 131;
         #statRecordLen := 72;
       ELSE
         RETURN; // No data set selected, abort execution
       END_IF;

       IF #readWrite = #MODE_WRITE THEN
         REGION write
           IF #appSpecificName THEN
             #statAppSpecName := #data.appSpecificName; // copy text into writing data
             #tempLen := LEN(#statAppSpecName); // determine length of text

             // Shift chars in array to remove String header
             FOR #tempIndex := 0 TO #tempLen - 1 DO
               #statRecord[#tempIndex] := #statRecord[#tempIndex + 2];
             END_FOR;

             // Fill remaining characters with null
             FOR #tempIndex := #tempLen TO #statRecordLen - 1 DO
               #statRecord[#tempIndex] := CHAR_TO_BYTE('$00');
             END_FOR;
           ELSIF #parameters THEN
             #statParameters := #data.parameters;
           ELSE // All other data sets are read only
             ;
           END_IF;
         END_REGION

       END_IF;
     END_IF;
   END_REGION

   REGION CALL
     #instDevice(execute     := #execute,
                 logicalAddr := #logicalAddr,
                 cap         := #cap,
                 readWrite   := #readWrite,
                 "port"      := #port,
                 index       := #statIndex,
                 subindex    := #statSubindex,
                 writeLen    := #statRecordLen,
                 timeout     := T#20s,
                 record      := #statRecord);
   END_REGION

   REGION READ
     // Copy data if available and valid
     IF #instDevice.done = TRUE AND #statDoneOld = FALSE AND #readWrite = #MODE_READ THEN
       IF #parameterPage0 THEN
         #data.parameterPage0 := #statParameterPage0;
       ELSIF #vendorName THEN
         #data.vendorName := #statVendorName;
       ELSIF #vendorText THEN
         #data.vendorText := #statVendorText;
       ELSIF #productName THEN
         #data.productName := #statProductName;
       ELSIF #productID THEN
         #data.productID := #statProductID;
       ELSIF #fwRevision THEN
         #data.firmwareRevision := #statFWRevision;
       ELSIF #appSpecificName THEN
         // Shift chars in array to make space for max/current length of String
         FOR #tempIndex := (#statRecordLen + 1) TO 2 BY -1 DO
           #statRecord[#tempIndex] := #statRecord[#tempIndex - 2];
         END_FOR;

         #statRecord[0] := INT_TO_BYTE(#statRecordLen); // manipulate array values for String 
         #statRecord[1] := INT_TO_BYTE(#statRecordLen);

         #data.appSpecificName := #statAppSpecName;
       ELSIF #diagnostics THEN
         #data.diagnostics := #statDiagnostics;
       ELSIF #measuredValues THEN
         #data.measuredValues := #statMeasuredValues;
       ELSIF #parameters THEN
         #data.parameters := #statParameters;
       ELSE // Other data sets are not defined
         ;
       END_IF;
     END_IF;

     #statDoneOld := #instDevice.done;
   END_REGION

   REGION OUTPUTS
     #done := #instDevice.done;
     #busy := #instDevice.busy;
     #error := #instDevice.error;
     #status := #instDevice.status;
     #diagDeviceFB := #instDevice.diagnostics;
   END_REGION
END_FUNCTION_BLOCK

FUNCTION_BLOCK "LIOLink_3SU1_IDKeySwitch"   // FB5210, SCL
TITLE = LIOLink_3SU1_IDKeySwitch / IO_LINK_3SU1_Keyswitch
{ S7_Optimized_Access := 'FALSE' }
AUTHOR : SIOS
FAMILY : LIOLink
VERSION : 2.0
// IO-Link Device FB for SIRIUS ACT ID Key Switch to use with S7-300/400 controllers! / IO-Link Geraete FB fuer SIRIUS 3SU1 ID-Schluesselschalter zur Nutzung mit S7-1500!
   VAR_INPUT
      execute : Bool;   // Request to execute function / Auftrag starten (mit steigender Flanke)
      logicalAddr : DInt;   // Logical address of IO-Link master module (sub module for ET 200eco PN) / Logische EA-Adresse des IO-Link Master Moduls
      cap : Int := 227;   // Client Access Point; 0xB400 for ET 200eco PN, CM 8x IO-Link, else 0xE003 (227) / Client Access Point (CAP), Siemens IO-Link Master immer 227 dezimal
      readWrite : Bool;   // FALSE: read, TRUE: write / Lese-/Schreibzugriff: 0=Lesen, 1=Schreiben
      port : Int;   // Port of the IO-Link Master for the Device / Port des Geraetes am IO-Link Mastermodul
      parameterPage0 : Bool;   // Read access on parameter page 0 / Lesen Parameter Page 0
      systemCommands : Bool;   // Write system commands / Write System Command to Switch
      vendorName : Bool;   // Read Vendor Name / Lesen Herstellername
      vendorText : Bool;   // Read Vendor Text / Lesen Herstellertext
      productName : Bool;   // Read Product Name / Lesen Produktname
      productID : Bool;   // Read Product ID / Lesen Produkt ID
      fwRevision : Bool;   // Read firmware revision / Lesen FW-Revision
      appSpecificName : Bool;   // Read/Write Application Specific Name / Lesen/Schreiben des spezifischen Applikationsnamen
      delKeyID : Bool;   // Read/Write: Delete key ID / Read / Write: Delete Key-ID
      keyList1 : Bool;   // Read keys 1 to key 30 / Read Key-List of Key 1 to Key 30
      keyList2 : Bool;   // Read keys 31 to key 50 / Read Key-List of Key 31 to Key 50
      diagnostics : Bool;   // Read diagnostics / Lesen der Gruppendiagnose
      insertedIDKey : Bool;   // Read ID of the inserted ID key / Read ID of the Currenty Key
      parameters : Bool;   // Read/write Parameters / Lesen/Schreiben der Parameter
   END_VAR
   VAR_OUTPUT
      done : Bool;   // TRUE: Commanded functionality has been completed successfully / Gueltigkeit 0: Daten ungueltig ; 1: Daten gueltig
      busy : Bool;   // TRUE: FB is not finished and new output values can be expected / 0: Auftrag beendet 1: Auftrag in Bearbeitung
      error : Bool;   // TRUE: An error occurred during the execution of the FB / Fehler = 0: kein Fehler; 1: Funktionsabbruch mit Fehler
      status : Word;   // 16#0000 - 16#7FFF: Status of the FB, 16#8000 - 16#FFFF: Error identification / DP/ PNIO - Fehlerstatus ; ERROR = 1 - Kommunikationsfehler in Detail
      diagDeviceFB : "LIOLink_typeDiagnostics";   // Diagnostics information of LIOLink_Device / IO-Link - Fehlerstatus; ERROR = 1: IO-Link Fehler in Detail
   END_VAR
   VAR_IN_OUT
      data : "LIOLink_3SU1_IDKeySwitch_typeAll";   // Data area, device specific (Data Type) / Ablage der Gerätedaten, gerätespezifisch (Datentyp in DB)
   END_VAR
   VAR
      instDevice : "LIOLink_Device";
      statRecordParam : Struct   // Parameters to read/write specific records / Datensatzparameter (geraetespezifisch)
         index : Array[0..28] of Int;   // Index of data set / Datensatzindex
         subindex : Array[0..28] of Int;   // Subindex of data sets / Datensatzsubindex
         length : Array[0..28] of Int;   // Length of data set / Datensatzlänge
      END_STRUCT;
      statRecord : Array[0..231] of Byte;   // Record buffer
      statParameterPage0 AT statRecord : "LIOLink_typeParameterPage0";
      statVendorName AT statRecord : String[10];
      statVendorText AT statRecord : String[64];
      statProductName AT statRecord : String[55];
      statProductID AT statRecord : String[18];
      statFWRevision AT statRecord : String[5];
      statAppSpecName AT statRecord : String[32];
      statDiagnostics AT statRecord : "LIOLink_3SU1_IDKeySwitch_typeDiag";
      statKeyList2 AT statRecord : "LIOLink_3SU1_IDKeySwitch_typeKeyList2";
      statKeyList1 AT statRecord : "LIOLink_3SU1_IDKeySwitch_typeKeyList1";
      statParameters AT statRecord : "LIOLink_3SU1_IDKeySwitch_typeParam";
      statInsertedKey AT statRecord : "LIOLink_3SU1_IDKeySwitch_typeInsertedKey";
      statDelKeyID AT statRecord : "LIOLink_3SU1_IDKeySwitch_typeKey";
      statSystemCommand AT statRecord : Byte;
      statIndex : Int;   // Requested index
      statSubindex : Int;   // Requested subindex
      statRecordLen : Int;   // Length of record to be written
      statRequest : Int;   // Case of request (data set) / Aktueller Fall (anfgefragter Datensatz)
      statDoneOld : Bool;   // Last cycle's value of instDevice.done
   END_VAR
   VAR_TEMP
      tempIndex : Int;   // Loop index
      tempLen : Int;   // Length
   END_VAR
   VAR CONSTANT
      MODE_READ : Bool := FALSE;   // Mode to read data
      MODE_WRITE : Bool := TRUE;   // Mode to write data
      STATUS_IDLE : Word := 16#7000;   // Status: Idle
   END_VAR
   // statRecordParam.index[4] := 0;
   // statRecordParam.index[3] := 0;
   // statRecordParam.index[2] := 2;
   // statRecordParam.index[1] := 0;
   // statRecordParam.index[24] := 0;
   // statRecordParam.index[23] := 92;
   // statRecordParam.index[21] := 82;
   // statRecordParam.index[20] := 81;
   // statRecordParam.index[19] := 80;
   // statRecordParam.index[18] := 24;
   // statRecordParam.index[17] := 23;
   // statRecordParam.index[16] := 22;
   // statRecordParam.index[15] := 21;
   // statRecordParam.index[14] := 20;
   // statRecordParam.index[13] := 19;
   // statRecordParam.index[12] := 18;
   // statRecordParam.index[11] := 17;
   // statRecordParam.index[10] := 16;
   // statRecordParam.index[8] := 0;
   // statRecordParam.index[7] := 0;
   // statRecordParam.index[6] := 0;
   // statRecordParam.index[5] := 0;
   // statRecordParam.length[28] := 0;
   // statRecordParam.length[27] := 20;
   // statRecordParam.length[26] := 22;
   // statRecordParam.length[25] := 0;
   // statRecordParam.length[24] := 0;
   // statRecordParam.length[23] := 20;
   // statRecordParam.length[22] := 0;
   // statRecordParam.length[21] := 120;
   // statRecordParam.length[20] := 180;
   // statRecordParam.length[19] := 5;
   // statRecordParam.length[18] := 32;
   // statRecordParam.length[17] := 5;
   // statRecordParam.length[16] := 5;
   // statRecordParam.length[15] := 8;
   // statRecordParam.length[13] := 18;
   // statRecordParam.length[12] := 55;
   // statRecordParam.length[11] := 64;
   // statRecordParam.length[10] := 10;
   // statRecordParam.length[9] := 0;
   // statRecordParam.length[8] := 0;
   // statRecordParam.length[7] := 0;
   // statRecordParam.length[6] := 0;
   // statRecordParam.length[5] := 0;
   // statRecordParam.length[4] := 0;
   // statRecordParam.length[3] := 0;
   // statRecordParam.length[2] := 1;
   // statRecordParam.length[1] := 16;
   // statRecordParam.length[0] := 0;
   // statRecordParam.index[28] := 0;
   // statRecordParam.index[27] := 131;
   // statRecordParam.index[26] := 94;
   // statRecordParam.index[25] := 0;
BEGIN
   REGION BLOCK INFO HEADER
     //===============================================================================
     // Siemens / (c)Copyright 2020
     //-------------------------------------------------------------------------------
     // Title:            LIOLink_3SU1_IDKeySwitch
     // Function:         Capsule block to communicate with 3SU1 ID Key Switch
     // Library:          LIOLink
     // Author:           Siemens Industry Online Support
     // Tested with:      CPU 317-2 PN/DP FW 3.2
     // Engineering:      TIA Portal V16
     // Restrictions:     --
     // Requirements:     --
     //-------------------------------------------------------------------------------
     // Change log table:
     // Version  | Date       | Expert in charge       | Changes applied
     //----------|------------|------------------------|------------------------------
     // 01.00.00 | 23.10.2015 | Online Support         | First release
     // 02.00.00 | 22.09.2020 | Online Support         | Rewrote block for FB "LIOLink_Device" V4.0.0
     //===============================================================================
   END_REGION

   REGION INIT
     IF (#execute = TRUE AND #instDevice.status = #STATUS_IDLE) THEN
       // Request selector
       IF #parameterPage0 THEN
         #statRequest := 1;
       ELSIF #systemCommands THEN
         #statRequest := 2;
       ELSIF #vendorName THEN
         #statRequest := 10;
       ELSIF #vendorText THEN
         #statRequest := 11;
       ELSIF #productName THEN
         #statRequest := 12;
       ELSIF #productID THEN
         #statRequest := 13;
       ELSIF #fwRevision THEN
         #statRequest := 17;
       ELSIF #appSpecificName THEN
         #statRequest := 18;
       ELSIF #delKeyID THEN
         #statRequest := 19;
       ELSIF #keyList1 THEN
         #statRequest := 20;
       ELSIF #keyList2 THEN
         #statRequest := 21;
       ELSIF #diagnostics THEN
         #statRequest := 23;
       ELSIF #insertedIDKey THEN
         #statRequest := 26;
       ELSIF #parameters THEN
         #statRequest := 27;
       ELSE
         #statRequest := 0;
       END_IF;

       // Set request specific parameters
       #statIndex := #statRecordParam.index[#statRequest];
       #statSubindex := #statRecordParam.subindex[#statRequest];
       #statRecordLen := #statRecordParam.length[#statRequest];

       IF #readWrite = #MODE_WRITE THEN
         REGION write
           CASE #statRequest OF
             1:
               #statParameterPage0 := #data.parameterPage0;
             2:
               #statSystemCommand := #data.systemCommand;
             18:
               #statAppSpecName := #data.appSpecificName; // copy text into writing data
               #tempLen := LEN(#statAppSpecName); // determine length of text

               // Shift chars in array to remove String header
               FOR #tempIndex := 0 TO #tempLen - 1 DO
                 #statRecord[#tempIndex] := #statRecord[#tempIndex + 2]; // move [2] to [0], [3] to [1] ... until end of String
               END_FOR;

               // Fill remaining characters with null
               FOR #tempIndex := #tempLen TO #statRecordLen - 1 DO
                 #statRecord[#tempIndex] := CHAR_TO_BYTE('$00');
               END_FOR;
             27:
               #statParameters := #data.parameters;
             ELSE // All other data sets are read only  
               ;
           END_CASE;
         END_REGION

       END_IF;
     END_IF;
   END_REGION

   REGION CALL
     #instDevice(execute     := #execute,
                 logicalAddr := #logicalAddr,
                 cap         := #cap,
                 readWrite   := #readWrite,
                 "port"      := #port,
                 index       := #statIndex,
                 subindex    := #statSubindex,
                 writeLen    := #statRecordLen,
                 timeout     := T#20s,
                 record      := #statRecord);
   END_REGION

   REGION READ
     // Copy data
     IF #instDevice.done = TRUE AND #statDoneOld = FALSE AND #readWrite = #MODE_READ THEN
       IF (#statRequest >= 10 AND #statRequest <= 18) THEN // Only applies for String parameters (case 10..18)
         // Shift all characters to add string header
         FOR #tempIndex := (#statRecordLen + 1) TO 2 BY -1 DO
           #statRecord[#tempIndex] := #statRecord[#tempIndex - 2];
         END_FOR;
         // Add String header
         #statRecord[0] := INT_TO_BYTE(#statRecordLen);
         #statRecord[1] := INT_TO_BYTE(#statRecordLen);
       END_IF;

       CASE #statRequest OF
         1:
           #data.parameterPage0 := #statParameterPage0;
         2:
           #data.systemCommand := #statSystemCommand;
         10:
           #data.vendorName := #statVendorName;
         11:
           #data.vendorText := #statVendorText;
         12:
           #data.productName := #statProductName;
         13:
           #data.productID := #statProductID;
         17:
           #data.fwRevision := #statFWRevision;
         18:
           #data.appSpecificName := #statAppSpecName;
         19:
           #data.delKeyID := #statDelKeyID;
         20:
           #data.keyList1 := #statKeyList1;
         21:
           #data.keyList2 := #statKeyList2;
         23:
           #data.diagnostics := #statDiagnostics;
         26:
           #data.insertedKey := #statInsertedKey;
         27:
           #data.parameters := #statParameters;
         ELSE // Other data sets are not defined
           ;
       END_CASE;
     END_IF;

     #statDoneOld := #instDevice.done;
   END_REGION

   REGION OUTPUTS
     #done := #instDevice.done;
     #busy := #instDevice.busy;
     #error := #instDevice.error;
     #status := #instDevice.status;
     #diagDeviceFB := #instDevice.diagnostics;
   END_REGION
END_FUNCTION_BLOCK

FUNCTION_BLOCK "LIOLink_3SU1_ElecModule"   // FB5220, SCL
TITLE = LIOLink_3SU1_ElecModule / IO_LINK_3SU1_Electronic
{ S7_Optimized_Access := 'FALSE' }
AUTHOR : SIOS
FAMILY : LIOLink
VERSION : 2.0
// IO-Link Device FB for SIRIUS ACT 3SU1 Electronic Module to use with S7-1200/1500 controllers! / IO-Link Geraete FB fuer SIRIUS 3SU1 Electronic Module zur Nutzung mit S7-1500!
   VAR_INPUT
      execute : Bool;   // Request to execute function / Auftrag starten (mit steigender Flanke)
      logicalAddr : DInt;   // Logical address of IO-Link master module (sub module for ET 200eco PN) / Logische EA-Adresse des IO-Link Master Moduls
      cap : Int := 227;   // Client Access Point; 0xB400 for ET 200eco PN, CM 8x IO-Link, else 0xE003 (227) / Client Access Point (CAP), Siemens IO-Link Master immer 227 dezimal
      readWrite : Bool;   // FALSE: read, TRUE: write / Lese-/Schreibzugriff: 0=Lesen, 1=Schreiben
      port : Int;   // Port of the IO-Link Master for the Device / Port des Geraetes am IO-Link Mastermodul
      parameterPage0 : Bool;   // Read access on parameter page 0 / Lesen Parameter Page 0
      systemCommand : Bool;   // Write System Command to Switch
      vendorName : Bool;   // Read Vendor Name / Lesen Herstellername
      vendorText : Bool;   // Read Vendor Text / Lesen Herstellertext
      productName : Bool;   // Read Product Name / Lesen Produktname
      productID : Bool;   // Read Product ID / Lesen Produkt ID
      fwRevision : Bool;   // Read FW-Revision / Lesen FW-Revision
      applicationSpecificName : Bool;   // Read/Write Application Specific Name / Lesen/Schreiben des spezifischen Applikationsnamen
      diagnostics : Bool;   // Read diagnostics / Lesen der Diagnose
      statistics : Bool;   // Read statistic data / Lesen der statistischen Daten
      parameters : Bool;   // Read / write Parameters / Lesen/Schreiben der Parameter
   END_VAR
   VAR_OUTPUT
      done : Bool;   // TRUE: Commanded functionality has been completed successfully / Gueltigkeit 0: Daten ungueltig ; 1: Daten gueltig
      busy : Bool;   // TRUE: FB is not finished and new output values can be expected / 0: Auftrag beendet 1: Auftrag in Bearbeitung
      error : Bool;   // TRUE: An error occurred during the execution of the FB / Fehler = 0: kein Fehler; 1: Funktionsabbruch mit Fehler
      status : Word;   // 16#0000 - 16#7FFF: Status of the FB, 16#8000 - 16#FFFF: Error identification / DP/ PNIO - Fehlerstatus ; ERROR = 1 - Kommunikationsfehler in Detail
      diagDeviceFB : "LIOLink_typeDiagnostics";   // Diagnostics information of LIOLink_Device / IO-Link - Fehlerstatus; ERROR = 1: IO-Link Fehler in Detail
   END_VAR
   VAR_IN_OUT
      data : "LIOLink_3SU1_ElecModule_typeAll";   // Data area, device specific (Data Type) / Ablage der Gerätedaten, gerätespezifisch (Datentyp in DB)
   END_VAR
   VAR
      instDevice : "LIOLink_Device";
      statRecordParam : Struct   // Parameters to read/write specific records / Datensatzparameter (geraetespezifisch)
         index : Array[0..28] of Int;   // Index of data set / Datensatzindex
         subindex : Array[0..28] of Int;   // Subindex of data sets / Datensatzsubindex
         length : Array[0..28] of Int;   // Length of data set / Datensatzlänge
      END_STRUCT;
      statRecord : Array[0..231] of Byte;   // Record buffer
      statParameterPage0 AT statRecord : "LIOLink_typeParameterPage0";
      statVendorName AT statRecord : String[10];
      statVendorText AT statRecord : String[58];
      statProductName AT statRecord : String[30];
      statProductID AT statRecord : String[8];
      statProductText AT statRecord : String[2];
      statSerialNumber AT statRecord : String[8];
      statHWRevision AT statRecord : String[4];
      statFWRevision AT statRecord : String[4];
      statAppSpecName AT statRecord : String[32];
      statDiagnostics AT statRecord : "LIOLink_3SU1_ElecModule_typeDiag";
      statParameters AT statRecord : "LIOLink_3SU1_ElecModule_typeParam";
      statSystemCommand AT statRecord : Byte;
      statStatistics AT statRecord : "LIOLink_3SU1_ElecModule_typeStats";
      statIndex : Int;   // Requested index
      statSubindex : Int;   // Requested subindex
      statRecordLen : Int;   // Length of record to be written
      statRequest : Int;   // Case of request (data set) / Aktueller Fall (anfgefragter Datensatz)
      statDone : Bool;   // Last cycle's value of instDevice.done
   END_VAR
   VAR_TEMP
      tempIndex : Int;   // Loop index
      tempLen : Int;   // Length
   END_VAR
   VAR CONSTANT
      MODE_READ : Bool := FALSE;   // Mode to read data
      MODE_WRITE : Bool := TRUE;   // Mode to write data
      STATUS_IDLE : Word := 16#7000;   // Status: Idle
   END_VAR
   // statRecordParam.index[1] := 0;
   // statRecordParam.index[2] := 2;
   // statRecordParam.index[3] := 0;
   // statRecordParam.index[4] := 0;
   // statRecordParam.index[5] := 0;
   // statRecordParam.index[6] := 0;
   // statRecordParam.index[7] := 0;
   // statRecordParam.index[8] := 0;
   // statRecordParam.index[10] := 16;
   // statRecordParam.index[11] := 17;
   // statRecordParam.index[12] := 18;
   // statRecordParam.index[13] := 19;
   // statRecordParam.index[14] := 20;
   // statRecordParam.index[15] := 21;
   // statRecordParam.index[16] := 22;
   // statRecordParam.index[17] := 23;
   // statRecordParam.index[18] := 24;
   // statRecordParam.index[19] := 80;
   // statRecordParam.index[20] := 94;
   // statRecordParam.index[21] := 100;
   // statRecordParam.index[23] := 92;
   // statRecordParam.index[24] := 0;
   // statRecordParam.index[25] := 0;
   // statRecordParam.index[27] := 131;
   // statRecordParam.index[28] := 0;
   // statRecordParam.length[0] := 0;
   // statRecordParam.length[1] := 16;
   // statRecordParam.length[2] := 1;
   // statRecordParam.length[3] := 0;
   // statRecordParam.length[4] := 0;
   // statRecordParam.length[5] := 0;
   // statRecordParam.length[6] := 0;
   // statRecordParam.length[7] := 0;
   // statRecordParam.length[8] := 0;
   // statRecordParam.length[9] := 0;
   // statRecordParam.length[10] := 10;
   // statRecordParam.length[11] := 64;
   // statRecordParam.length[12] := 55;
   // statRecordParam.length[13] := 18;
   // statRecordParam.length[15] := 16;
   // statRecordParam.length[16] := 6;
   // statRecordParam.length[17] := 6;
   // statRecordParam.length[18] := 32;
   // statRecordParam.length[19] := 5;
   // statRecordParam.length[20] := 48;
   // statRecordParam.length[21] := 0;
   // statRecordParam.length[22] := 0;
   // statRecordParam.length[23] := 23;
   // statRecordParam.length[24] := 0;
   // statRecordParam.length[25] := 0;
   // statRecordParam.length[26] := 43;
   // statRecordParam.length[27] := 126;
   // statRecordParam.length[28] := 0;
BEGIN
   REGION BLOCK INFO HEADER
     //===============================================================================
     // Siemens / (c)Copyright 2020
     //-------------------------------------------------------------------------------
     // Title:            LIOLink_3SU1_ElecModule
     // Function:         Capsule block to communicate with 3SU1 Electronic Module
     // Library:          LIOLink
     // Author:           Siemens Industry Online Support
     // Tested with:      CPU 317-2 PN/DP FW 3.2
     // Engineering:      TIA Portal V16
     // Restrictions:     --
     // Requirements:     --
     //-------------------------------------------------------------------------------
     // Change log table:
     // Version  | Date       | Expert in charge       | Changes applied
     //----------|------------|------------------------|------------------------------
     // 01.00.00 | 23.10.2015 | Online Support         | First release
     // 02.00.00 | 22.09.2020 | Online Support         | Rewrote block for FB "LIOLink_Device" V4.0.0
     //===============================================================================
   END_REGION

   REGION INIT
     IF (#execute = TRUE AND #instDevice.busy = FALSE) THEN
       // Request selector
       IF #parameterPage0 THEN
         #statRequest := 1;
       ELSIF #systemCommand THEN
         #statRequest := 2;
       ELSIF #vendorName THEN
         #statRequest := 10;
       ELSIF #vendorText THEN
         #statRequest := 11;
       ELSIF #productName THEN
         #statRequest := 12;
       ELSIF #productID THEN
         #statRequest := 13;
       ELSIF #fwRevision THEN
         #statRequest := 17;
       ELSIF #applicationSpecificName THEN
         #statRequest := 18;
       ELSIF #statistics THEN
         #statRequest := 20;
       ELSIF #diagnostics THEN
         #statRequest := 23;
       ELSIF #parameters THEN
         #statRequest := 27;
       ELSE
         #statRequest := 0;
       END_IF;

       #statIndex := #statRecordParam.index[#statRequest];
       #statSubindex := #statRecordParam.subindex[#statRequest];
       #statRecordLen := #statRecordParam.length[#statRequest];

       IF #readWrite = #MODE_WRITE THEN
         REGION write
           CASE #statRequest OF
             1:
               #statParameterPage0 := #data.parameterPage0;
             2:
               #statSystemCommand := #data.systemCommand;
             18:
               #statAppSpecName := #data.appSpecificName; // copy text into writing data
               #tempLen := LEN(#statAppSpecName); // determine length of text

               // Shift chars in array to remove String header
               FOR #tempIndex := 0 TO #tempLen - 1 DO
                 #statRecord[#tempIndex] := #statRecord[#tempIndex + 2]; // move [2] to [0], [3] to [1] ... until end of String
               END_FOR;

               // Fill remaining characters
               FOR #tempIndex := #tempLen TO #statRecordLen - 1 DO
                 #statRecord[#tempIndex] := CHAR_TO_BYTE('$00');
               END_FOR;
             27:
               #statParameters := #data.parameters;
             ELSE    // all other data sets are read only  
               ;
           END_CASE;
         END_REGION

       END_IF;
     END_IF;
   END_REGION

   REGION CALL
     #instDevice(execute     := #execute,
                 logicalAddr := #logicalAddr,
                 cap         := #cap,
                 readWrite   := #readWrite,
                 "port"      := #port,
                 index       := #statIndex,
                 subindex    := #statSubindex,
                 writeLen    := #statRecordLen,
                 timeout     := T#20s,
                 record      := #statRecord);
   END_REGION

   REGION READ
     // Copy data if available and valid
     IF #instDevice.done = TRUE AND #statDone = FALSE AND #readWrite = #MODE_READ THEN
       IF (#statRequest >= 10 AND #statRequest <= 18) THEN // Only applies for STRING parameters (case 10..18)
         // add two to data set length for STRING parameters (max./current length)
         FOR #tempIndex := (#statRecordLen + 1) TO 2 BY -1 DO
           #statRecord[#tempIndex] := #statRecord[#tempIndex - 2];
         END_FOR; // Shift chars in array to make space for max/current length of STRING

         #statRecord[0] := INT_TO_BYTE(#statRecordLen); // manipulate array values for STRING 
         #statRecord[1] := INT_TO_BYTE(#statRecordLen);
       END_IF; // Shift all strings and add string header 

       CASE #statRequest OF
         1:
           #data.parameterPage0 := #statParameterPage0;
         2:
           #data.systemCommand := #statSystemCommand;
         10:
           #data.vendorName := #statVendorName;
         11:
           #data.vendorText := #statVendorText;
         12:
           #data.productName := #statProductName;
         13:
           #data.productID := #statProductID;
         17:
           #data.fwRevision := #statFWRevision;
         18:
           #data.appSpecificName := #statAppSpecName;
         20:
           #data.statistics := #statStatistics;
         23:
           #data.diagnostics := #statDiagnostics;
         27:
           #data.parameters := #statParameters;
         ELSE // all other data sets are not defined
           ;
       END_CASE;
     END_IF;

     #statDone := #instDevice.done;
   END_REGION

